	E_Element_State_Long.eWaterReady:;
			IF eReq=E_Request_List.eDissolve THEN;
				eProcess:=E_Element_Process.eDissolving;
			END_IF	
			IF eReq=E_Request_List.eFinish THEN;
				mClearProduction(state:=E_Element_State_Long.eStandby);
			END_IF
	E_Element_State_Long.eReady:;
			IF eReq=E_Request_List.eProduction THEN;
				eProcess:=E_Element_Process.eConnectionToLine;
			END_IF	
			IF eReq=E_Request_List.eFinish THEN;
				mClearProduction(state:=E_Element_State_Long.eStandby);
			END_IF			

	E_Element_State_Long.eProduction:;
			IF eReq=E_Request_List.eDisconnectTank THEN;
				eProcess:=E_Element_Process.eDisconnection;
			END_IF	
			
			IF fbInterConnection_ProL.bAvalableToDisconnect 
			AND m_Production_Run_Pump()
			THEN;
				IF memo_Production_Storage_Mode THEN;
					fb_PumpLine.m_Run(RPM:=stProdParam.stRecipe.FlowRate_Storage);
				ELSE;
					fb_PumpLine.m_Run(RPM:=stProdParam.stRecipe.FlowRate_Production);
				END_IF
				
			ELSE;
				fb_PumpLine.m_Stop();
			END_IF		

	E_Element_State_Long.eEmpty:;
			IF eReq=E_Request_List.eFinish THEN;
				mClearProduction(state:=E_Element_State_Long.eStandby);
			END_IF	

	E_Element_State_Long.eExpired:;
		CASE refElement.eState_Long_Expiered OF
			
			E_Element_State_Long.eProduction:;	
				IF eReq=E_Request_List.eDisconnectTank THEN;
					eProcess:=E_Element_Process.eDisconnection;
				END_IF
				
				IF fbInterConnection_ProL.bAvalableToDisconnect 
				AND m_Production_Run_Pump()
				THEN;
					IF memo_Production_Storage_Mode THEN;
						fb_PumpLine.m_Run(RPM:=stProdParam.stRecipe.FlowRate_Storage);
					ELSE;
						fb_PumpLine.m_Run(RPM:=stProdParam.stRecipe.FlowRate_Production);
					END_IF
					
				ELSE;
					fb_PumpLine.m_Stop();
				END_IF	
		ELSE
			IF eReq=E_Request_List.eFinish THEN;
				mClearProduction(state:=E_Element_State_Long.eStandby);
			END_IF			
		END_CASE
		
END_CASE
END_ACTION

ACTION _aReady_entry:

END_ACTION

ACTION _aReady_exit:
bRun:=TRUE;
bDone:=FALSE;
//bCntrlTemp:=TRUE;
END_ACTION

ACTION _aStart_TriPump_1_active:
bStepDone:=TRUE;
END_ACTION

ACTION _aStart_TriPump_1_entry:
fb_PumpTriBlender.m_Run(RPM:=stProdParam.stRecipe.FlowRate_WaterPushing);
END_ACTION

ACTION _aStart_TriPump_2_active:
bStepDone:=TRUE;
END_ACTION

ACTION _aStart_TriPump_2_entry:
fb_PumpTriBlender.m_Run(RPM:=stProdParam.stRecipe.FlowRate_WaterPushing);
END_ACTION

ACTION _aStart_TriPump_3_active:
bStepDone:=TRUE;
END_ACTION

ACTION _aStart_TriPump_3_entry:
fb_PumpTriBlender.m_Run(RPM:=stProdParam.stRecipe.FlowRate_WaterPushing);
memo_Tank_Level_start:=ref_fbTankSensors.act_Volume;
END_ACTION

ACTION _aState_Update_01_entry:
refState_Long:=E_Element_State_Long.eNotClean;
END_ACTION

ACTION _aState_Update_02_entry:
refState_Long:=E_Element_State_Long.eWaterReady;
END_ACTION

ACTION _aState_Update_03_entry:
refState_Long:=E_Element_State_Long.eReady;
END_ACTION

ACTION _aState_Update_04_entry:
refState_Long:=E_Element_State_Long.eProduction;
END_ACTION

ACTION _aState_Update_05_entry:
refState_Long:=E_Element_State_Long.eReady;
END_ACTION

ACTION _aStop_TriPump_1_active:
bStepDone:=TRUE;
END_ACTION

ACTION _aStop_TriPump_1_entry:
fb_PumpTriBlender.m_Stop();
END_ACTION

ACTION _aStop_TriPump_2_active:
bStepDone:=TRUE;
END_ACTION

ACTION _aStop_TriPump_2_entry:
fb_PumpTriBlender.m_Stop();
END_ACTION

ACTION _aStop_TriPump_3_active:
bStepDone:=TRUE;
END_ACTION

ACTION _aStop_TriPump_3_entry:
fb_PumpTriBlender.m_Stop();
END_ACTION

ACTION _aTank_Drain_active:
bStepDone:=FALSE;
IF fbTarget.m_CheckStatus(eReqStatus:=E_Tank_Target.eDrain) THEN;
	bTON_Active:=TRUE;
	
ELSIF Tank_Drain.t>=T#3S THEN; // max time to detect drain open
	bStepDone:=TRUE;
END_IF
IF Call_TON.Q THEN
	bStepDone:=TRUE;
END_IF
END_ACTION

ACTION _aTank_Drain_entry:
fbTarget.m_Run(eReqProc:=E_Tank_Target.eDrain);
bTON_Active:=FALSE;
END_ACTION

ACTION _aTank_Open_active:
bStepDone:=FALSE;
IF fbTarget.m_CheckStatus(eReqStatus:=E_Tank_Target.eOpen) THEN;
	bTON_Active:=TRUE;
END_IF
IF Call_TON.Q THEN
	bStepDone:=TRUE;
END_IF
END_ACTION

ACTION _aTank_Open_entry:
fbTarget.m_Run(eReqProc:=E_Tank_Target.eOpen);
bTON_Active:=FALSE;
END_ACTION

ACTION _aWater_Fill_active:
bStepDone:=FALSE;
IF TRUE 
AND TRUE//Reserved for tank level from recipe
//AND ref_fbTankSensors.get_stTankLevel().rTankLevel>=stProdParam.stRecipe.arr_Component[1].rWeight
AND fbTarget.stTankLevel.rTankLevel>=stProdParam.stRecipe.arr_Component[1].rWeight
THEN;
	bStepDone:=TRUE;
	
//temp overweight protection
ELSIF stT3_Sens.rTankLevel+stT4_Sens.rTankLevel>1000 THEN;
	bStepDone:=TRUE;
	
ELSIF bRunOffline 
AND Water_Fill.t>=T#10S
THEN
	bStepDone:=TRUE;
END_IF
END_ACTION

ACTION act_Call_Interface:
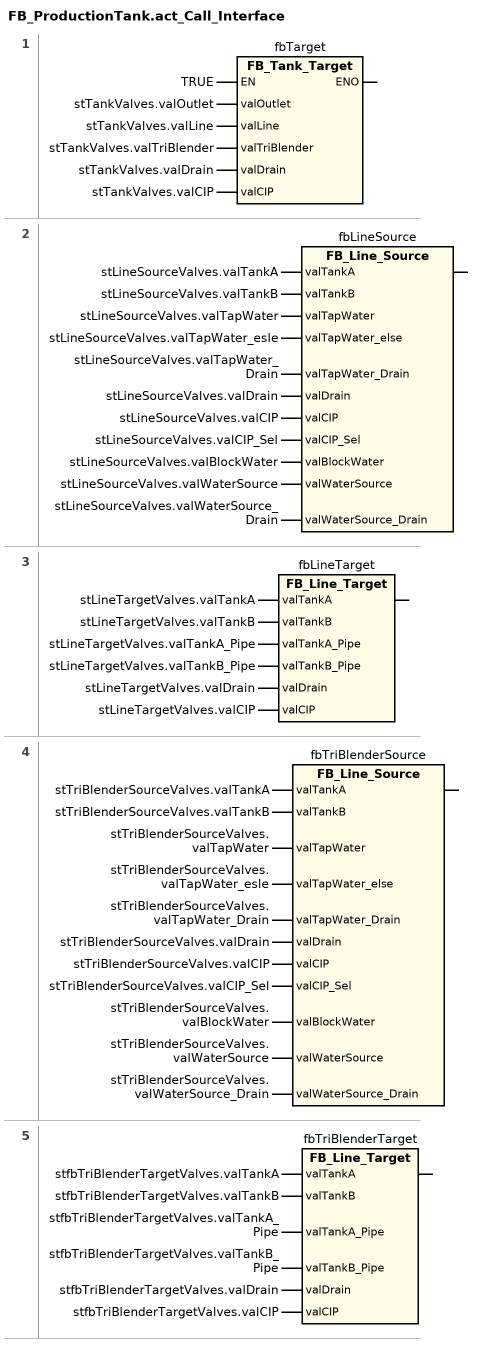
// NETWORK 1
fbTarget(
    valOutlet := stTankValves.valOutlet,
    valLine := stTankValves.valLine,
    valTriBlender := stTankValves.valTriBlender,
    valDrain := stTankValves.valDrain,
    valCIP := stTankValves.valCIP); // FB_Tank_Target

// NETWORK 2
fbLineSource(
    valTankA := stLineSourceValves.valTankA,
    valTankB := stLineSourceValves.valTankB,
    valTapWater := stLineSourceValves.valTapWater,
    valTapWater_else := stLineSourceValves.valTapWater_esle,
    valTapWater_Drain := stLineSourceValves.valTapWater_Drain,
    valDrain := stLineSourceValves.valDrain,
    valCIP := stLineSourceValves.valCIP,
    valCIP_Sel := stLineSourceValves.valCIP_Sel,
    valBlockWater := stLineSourceValves.valBlockWater,
    valWaterSource := stLineSourceValves.valWaterSource,
    valWaterSource_Drain := stLineSourceValves.valWaterSource_Drain); // FB_Line_Source

// NETWORK 3
fbLineTarget(
    valTankA := stLineTargetValves.valTankA,
    valTankB := stLineTargetValves.valTankB,
    valTankA_Pipe := stLineTargetValves.valTankA_Pipe,
    valTankB_Pipe := stLineTargetValves.valTankB_Pipe,
    valDrain := stLineTargetValves.valDrain,
    valCIP := stLineTargetValves.valCIP); // FB_Line_Target

// NETWORK 4
fbTriBlenderSource(
    valTankA := stTriBlenderSourceValves.valTankA,
    valTankB := stTriBlenderSourceValves.valTankB,
    valTapWater := stTriBlenderSourceValves.valTapWater,
    valTapWater_else := stTriBlenderSourceValves.valTapWater_esle,
    valTapWater_Drain := stTriBlenderSourceValves.valTapWater_Drain,
    valDrain := stTriBlenderSourceValves.valDrain,
    valCIP := stTriBlenderSourceValves.valCIP,
    valCIP_Sel := stTriBlenderSourceValves.valCIP_Sel,
    valBlockWater := stTriBlenderSourceValves.valBlockWater,
    valWaterSource := stTriBlenderSourceValves.valWaterSource,
    valWaterSource_Drain := stTriBlenderSourceValves.valWaterSource_Drain); // FB_Line_Source

// NETWORK 5
fbTriBlenderTarget(
    valTankA := stfbTriBlenderTargetValves.valTankA,
    valTankB := stfbTriBlenderTargetValves.valTankB,
    valTankA_Pipe := stfbTriBlenderTargetValves.valTankA_Pipe,
    valTankB_Pipe := stfbTriBlenderTargetValves.valTankB_Pipe,
    valDrain := stfbTriBlenderTargetValves.valDrain,
    valCIP := stfbTriBlenderTargetValves.valCIP); // FB_Line_Target

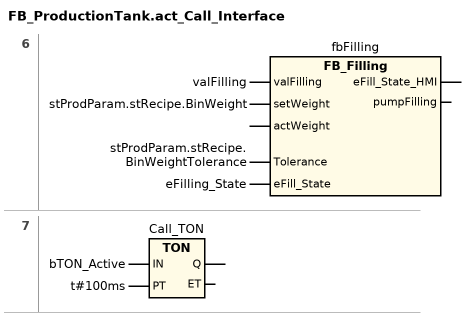
// NETWORK 6
fbFilling(
    valFilling := valFilling,
    setWeight := stProdParam.stRecipe.BinWeight,
    Tolerance := stProdParam.stRecipe.BinWeightTolerance,
    eFill_State := eFilling_State); // FB_Filling

// NETWORK 7
Call_TON(IN := bTON_Active, PT := t#100ms); // TON
END_ACTION

ACTION act_ExpirationTime:
IF stProdParam.eStatus=E_Prod_Status.Active 
THEN;
	refElement.m_Set_ExpirationDuration(eExTime_set:=E_ExTime.eProduct, setTime:=stProdParam.stRecipe.ExpirationTime);
	refElement.m_Set_ExpirationDuration(eExTime_set:=E_ExTime.eWater, setTime:=stProdParam.stRecipe.ExpirationTime_Water);
END_IF


(*
IF stProdParam.eStatus=E_Prod_Status.Active 
AND refElement.State>=E_Element_State_Long.eWaterReady
THEN;
	IF refElement.memoDissolving_active 
	//OR eStatus>=E_Element_State_Long.eReady
	THEN
		refElement.ExpirationTime:=stProdParam.stRecipe.ExpirationTime;
	ELSE;
		refElement.ExpirationTime:=stProdParam.stRecipe.ExpirationTime_Water;
	END_IF
	
ELSE;
	refElement.ExpirationTime:=ExDuration_Default;
END_IF
*)
END_ACTION

ACTION act_Filling:


IF TRUE 
AND bReady
AND refElement.eState_Long=E_Element_State_Long.eProduction
AND TRUE
AND TRUE
THEN;
	CASE pFilling_State OF 
		E_Filling_State.eNot_Ready:;
				pFilling_State:=E_Filling_State.eReady_ToFill;
				
		E_Filling_State.eReady_ToFill:;
				//
		E_Filling_State.eFilling_InProcess:;
				//
		
	END_CASE
ELSE;
	pFilling_State:=E_Filling_State.eNot_Ready;
END_IF

refElement.pFilling_State:=pFilling_State;

(*
IF fbInterConnection_ProL.bActive THEN;
	IF trn_Tank_Marinade THEN;
		fbElement[E_Element_List.eLine_Marinada].pFilling_State:=pFilling_State;
	ELSIF trn_Tank_Color THEN;
		fbElement[E_Element_List.eLine_Color].pFilling_State:=pFilling_State;
	END_IF	
END_IF
*)
END_ACTION

ACTION act_GetReference:
m_Set_SFCFlags_Reference();
refElement REF= fbElement[eElementID];
refState_Long REF= fbElement[eElementID].eState_Long;
//stPis_FillWater REF= stPis[valFillWater];
//stPis_FillWaterDrain REF= stPis[valFillWaterDrain];
//stPis_DrainTapWater REF= stPis[valDrainTapWater];

ref_fbTankSensors REF= g_Data.arrTanksSens[eTank_Name];
stTank_Level:=ref_fbTankSensors.get_stTankLevel();
fbTarget.set_TankLevel(set_stTankLevel:=stTank_Level);

stPis_CWIn REF= stPis[valCW_In];
stPis_CWOut	 REF= stPis[valCW_Out];

eStatus:=refState_Long;

//bRunCIP :=g_Data.b_CIP_Run;
bRunCIP := g_Data.fbElement[eElementID].m_Get_InterConnection() = E_InterConnection.ConnToCIP;
(*
stPis_Outlet		REF= g_Piston.stPis[valOutlet];
stPis_Line			REF= g_Piston.stPis[valOutlet];
stPis_TriBlender	REF= g_Piston.stPis[valOutlet];
stPis_Drain			REF= g_Piston.stPis[valOutlet];
stPis_CIP			REF= g_Piston.stPis[valOutlet];
*)
END_ACTION

ACTION act_Oper:
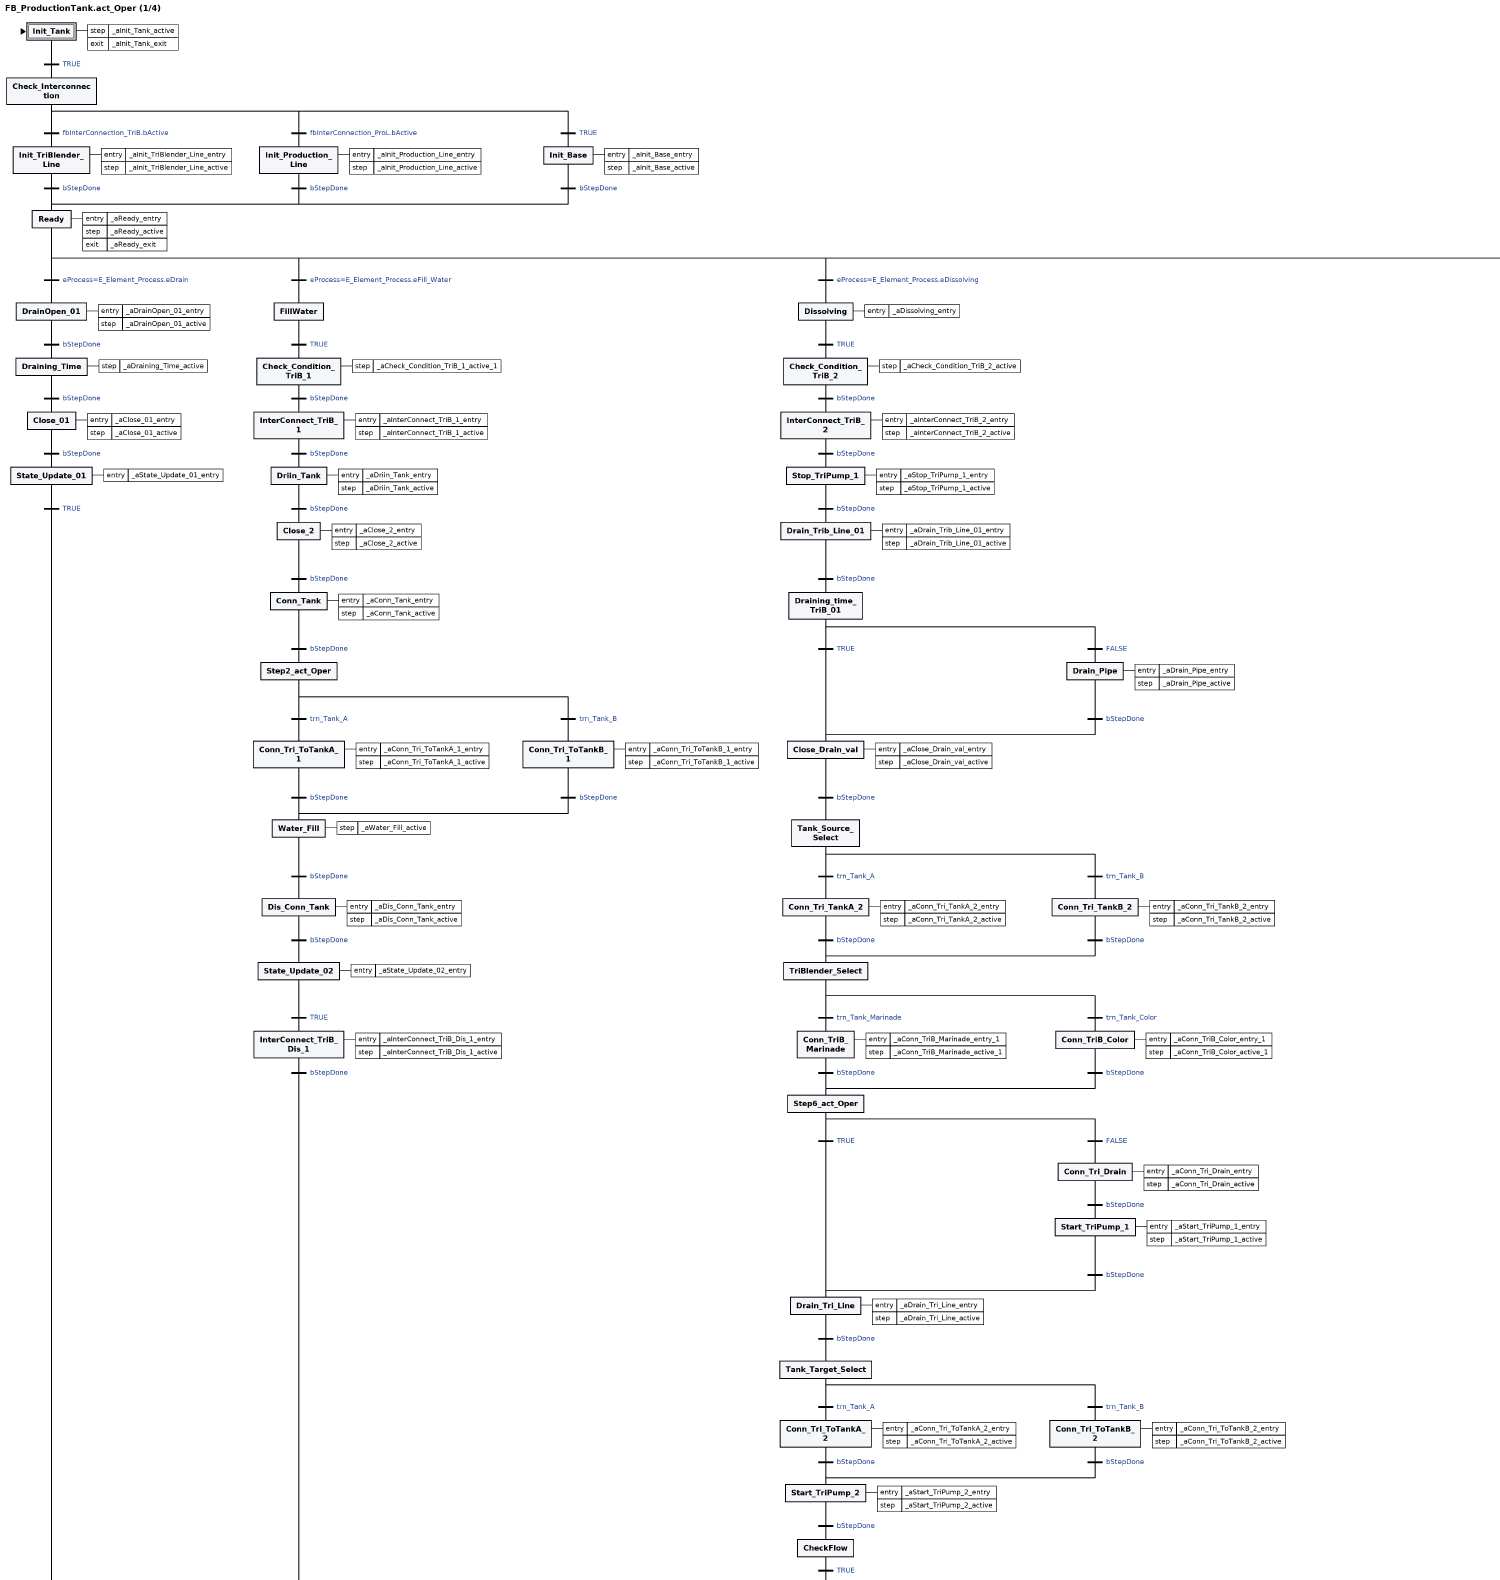
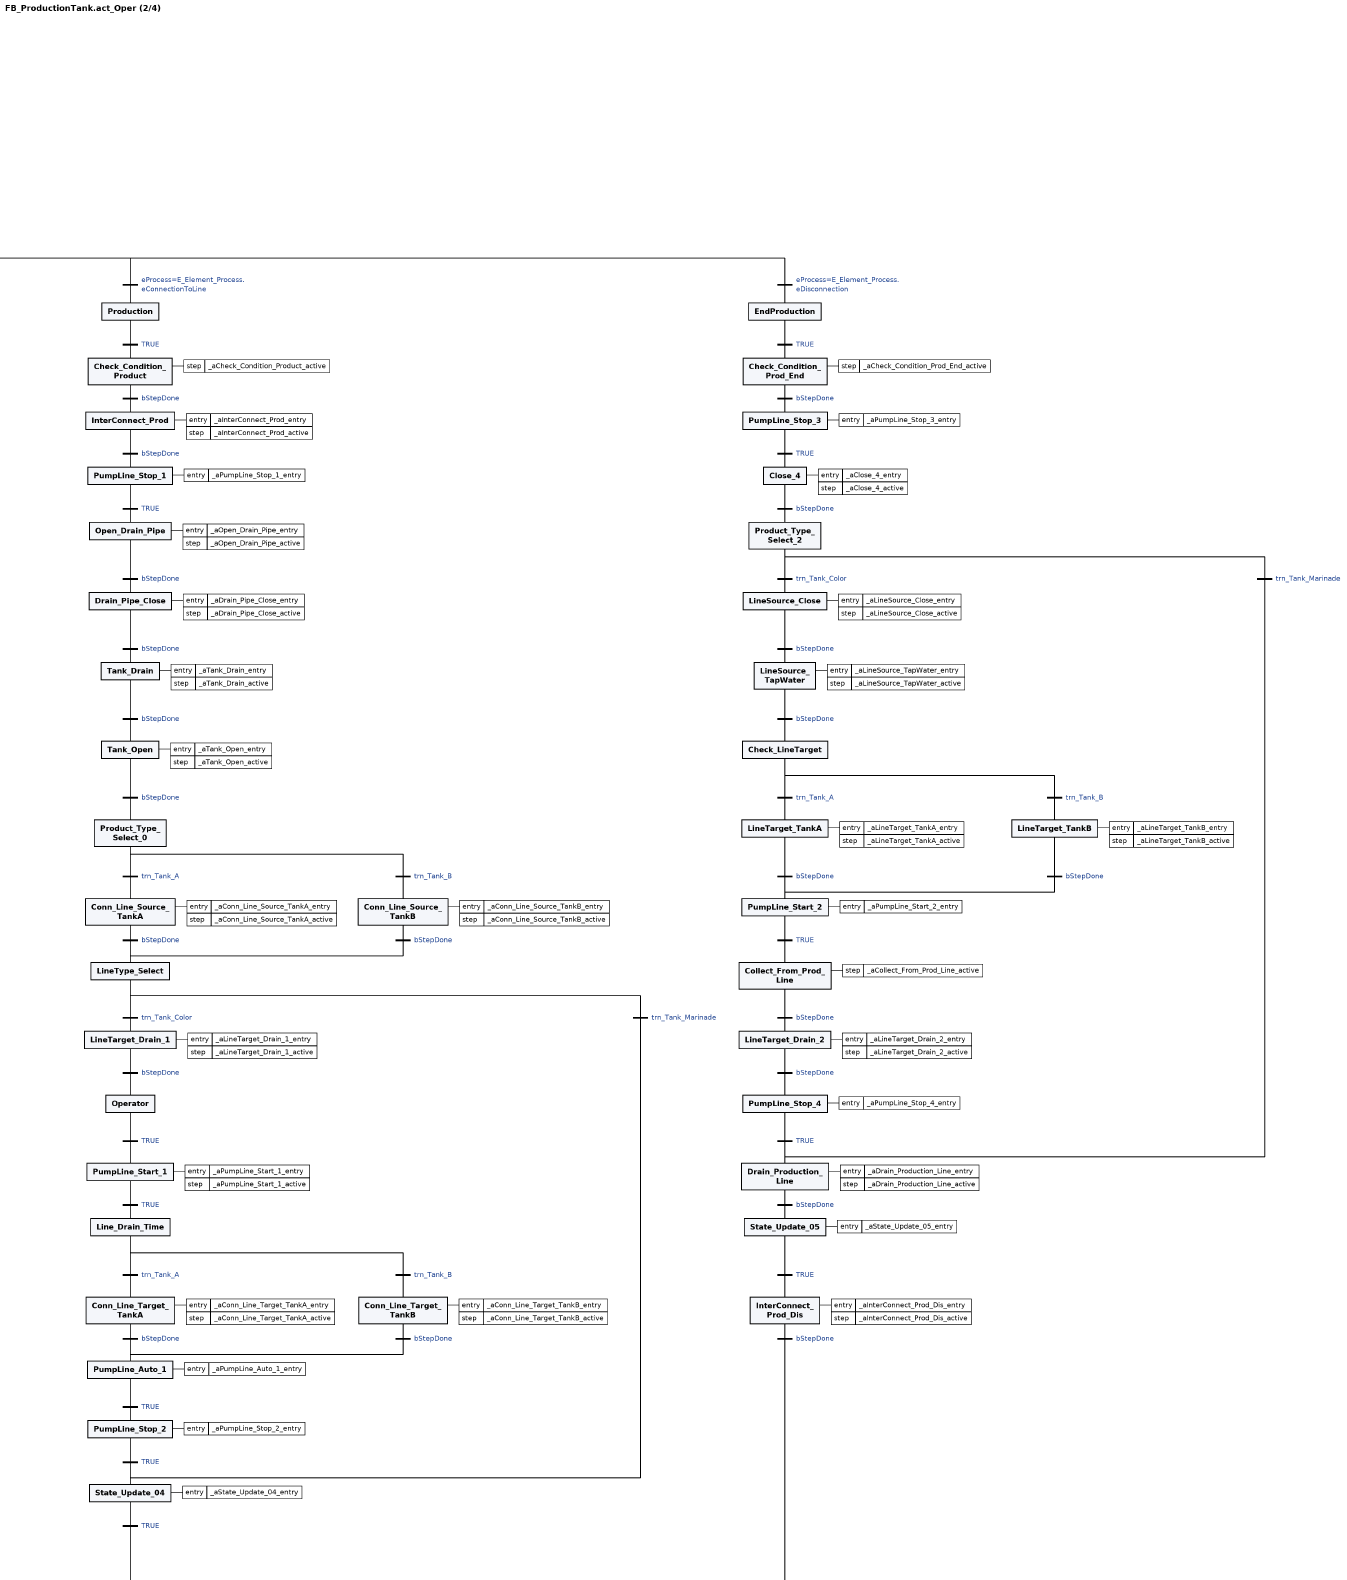
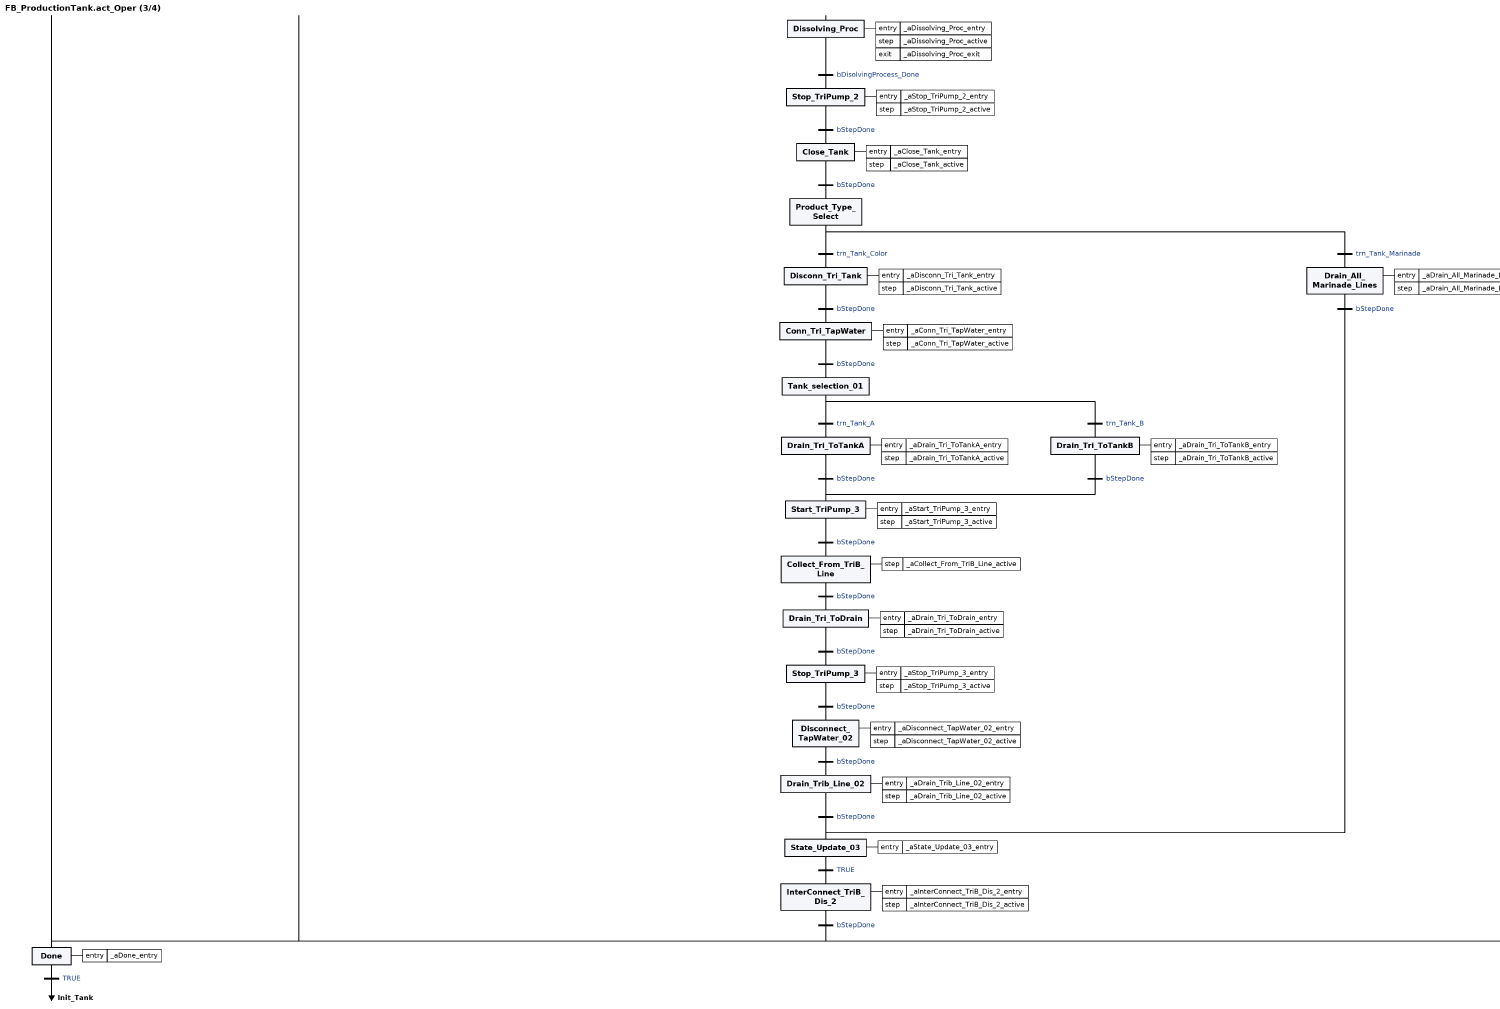
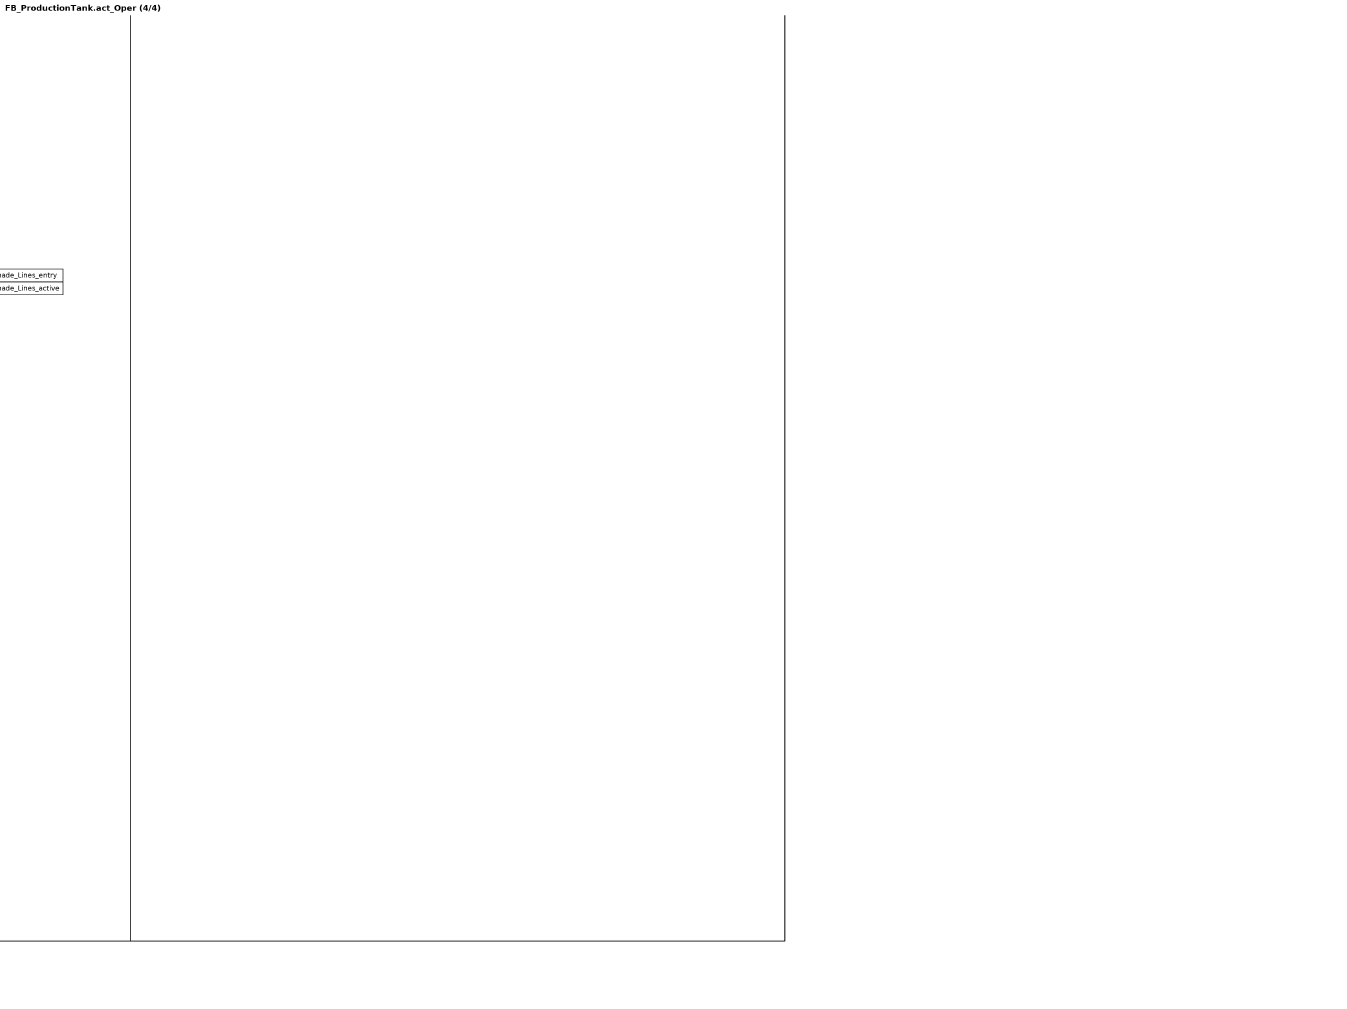
INITIAL_STEP Init_Tank:
    _aInit_Tank_active(N);  // step action
    _aInit_Tank_exit(P0);  // exit action
END_STEP
TRANSITION FROM Init_Tank TO Check_Interconnection
    := TRUE;
END_TRANSITION
STEP Check_Interconnection:
END_STEP
TRANSITION FROM Check_Interconnection TO Init_TriBlender_Line
    := fbInterConnection_TriB.bActive;
END_TRANSITION
STEP Init_TriBlender_Line:
    _aInit_TriBlender_Line_entry(P1);  // entry action
    _aInit_TriBlender_Line_active(N);  // step action
END_STEP
TRANSITION FROM Init_TriBlender_Line TO Ready
    := bStepDone;
END_TRANSITION
TRANSITION FROM Check_Interconnection TO Init_Production_Line
    := fbInterConnection_ProL.bActive;
END_TRANSITION
STEP Init_Production_Line:
    _aInit_Production_Line_entry(P1);  // entry action
    _aInit_Production_Line_active(N);  // step action
END_STEP
TRANSITION FROM Init_Production_Line TO Ready
    := bStepDone;
END_TRANSITION
TRANSITION FROM Check_Interconnection TO Init_Base
    := TRUE;
END_TRANSITION
STEP Init_Base:
    _aInit_Base_entry(P1);  // entry action
    _aInit_Base_active(N);  // step action
END_STEP
TRANSITION FROM Init_Base TO Ready
    := bStepDone;
END_TRANSITION
STEP Ready:
    _aReady_entry(P1);  // entry action
    _aReady_active(N);  // step action
    _aReady_exit(P0);  // exit action
END_STEP
TRANSITION FROM Ready TO DrainOpen_01
    := eProcess=E_Element_Process.eDrain;
END_TRANSITION
STEP DrainOpen_01:  // min time T#2s
    _aDrainOpen_01_entry(P1);  // entry action
    _aDrainOpen_01_active(N);  // step action
END_STEP
TRANSITION FROM DrainOpen_01 TO Draining_Time
    := bStepDone;
END_TRANSITION
STEP Draining_Time:  // min time T#2s
    _aDraining_Time_active(N);  // step action
END_STEP
TRANSITION FROM Draining_Time TO Close_01
    := bStepDone;
END_TRANSITION
STEP Close_01:  // min time T#2s
    _aClose_01_entry(P1);  // entry action
    _aClose_01_active(N);  // step action
END_STEP
TRANSITION FROM Close_01 TO State_Update_01
    := bStepDone;
END_TRANSITION
STEP State_Update_01:
    _aState_Update_01_entry(P1);  // entry action
END_STEP
TRANSITION FROM State_Update_01 TO Done
    := TRUE;
END_TRANSITION
TRANSITION FROM Ready TO FillWater
    := eProcess=E_Element_Process.eFill_Water;
END_TRANSITION
STEP FillWater:
END_STEP
TRANSITION FROM FillWater TO Check_Condition_TriB_1
    := TRUE;
END_TRANSITION
STEP Check_Condition_TriB_1:
    _aCheck_Condition_TriB_1_active_1(N);  // step action
END_STEP
TRANSITION FROM Check_Condition_TriB_1 TO InterConnect_TriB_1
    := bStepDone;
END_TRANSITION
STEP InterConnect_TriB_1:
    _aInterConnect_TriB_1_entry(P1);  // entry action
    _aInterConnect_TriB_1_active(N);  // step action
END_STEP
TRANSITION FROM InterConnect_TriB_1 TO Driin_Tank
    := bStepDone;
END_TRANSITION
STEP Driin_Tank:  // min time t#2s
    _aDriin_Tank_entry(P1);  // entry action
    _aDriin_Tank_active(N);  // step action
END_STEP
TRANSITION FROM Driin_Tank TO Close_2
    := bStepDone;
END_TRANSITION
STEP Close_2:  // min time t#2s
    _aClose_2_entry(P1);  // entry action
    _aClose_2_active(N);  // step action
END_STEP
TRANSITION FROM Close_2 TO Conn_Tank
    := bStepDone;
END_TRANSITION
STEP Conn_Tank:  // min time t#2s
    _aConn_Tank_entry(P1);  // entry action
    _aConn_Tank_active(N);  // step action
END_STEP
TRANSITION FROM Conn_Tank TO Step2_act_Oper
    := bStepDone;
END_TRANSITION
STEP Step2_act_Oper:
END_STEP
TRANSITION FROM Step2_act_Oper TO Conn_Tri_ToTankA_1
    := trn_Tank_A;
END_TRANSITION
STEP Conn_Tri_ToTankA_1:
    _aConn_Tri_ToTankA_1_entry(P1);  // entry action
    _aConn_Tri_ToTankA_1_active(N);  // step action
END_STEP
TRANSITION FROM Conn_Tri_ToTankA_1 TO Water_Fill
    := bStepDone;
END_TRANSITION
TRANSITION FROM Step2_act_Oper TO Conn_Tri_ToTankB_1
    := trn_Tank_B;
END_TRANSITION
STEP Conn_Tri_ToTankB_1:
    _aConn_Tri_ToTankB_1_entry(P1);  // entry action
    _aConn_Tri_ToTankB_1_active(N);  // step action
END_STEP
TRANSITION FROM Conn_Tri_ToTankB_1 TO Water_Fill
    := bStepDone;
END_TRANSITION
STEP Water_Fill:  // min time t#2s
    _aWater_Fill_active(N);  // step action
END_STEP
TRANSITION FROM Water_Fill TO Dis_Conn_Tank
    := bStepDone;
END_TRANSITION
STEP Dis_Conn_Tank:  // min time t#2s
    _aDis_Conn_Tank_entry(P1);  // entry action
    _aDis_Conn_Tank_active(N);  // step action
END_STEP
TRANSITION FROM Dis_Conn_Tank TO State_Update_02
    := bStepDone;
END_TRANSITION
STEP State_Update_02:  // min time t#2s
    _aState_Update_02_entry(P1);  // entry action
END_STEP
TRANSITION FROM State_Update_02 TO InterConnect_TriB_Dis_1
    := TRUE;
END_TRANSITION
STEP InterConnect_TriB_Dis_1:
    _aInterConnect_TriB_Dis_1_entry(P1);  // entry action
    _aInterConnect_TriB_Dis_1_active(N);  // step action
END_STEP
TRANSITION FROM InterConnect_TriB_Dis_1 TO Done
    := bStepDone;
END_TRANSITION
TRANSITION FROM Ready TO Dissolving
    := eProcess=E_Element_Process.eDissolving;
END_TRANSITION
STEP Dissolving:
    _aDissolving_entry(P1);  // entry action
END_STEP
TRANSITION FROM Dissolving TO Check_Condition_TriB_2
    := TRUE;
END_TRANSITION
STEP Check_Condition_TriB_2:
    _aCheck_Condition_TriB_2_active(N);  // step action
END_STEP
TRANSITION FROM Check_Condition_TriB_2 TO InterConnect_TriB_2
    := bStepDone;
END_TRANSITION
STEP InterConnect_TriB_2:
    _aInterConnect_TriB_2_entry(P1);  // entry action
    _aInterConnect_TriB_2_active(N);  // step action
END_STEP
TRANSITION FROM InterConnect_TriB_2 TO Stop_TriPump_1
    := bStepDone;
END_TRANSITION
STEP Stop_TriPump_1:
    _aStop_TriPump_1_entry(P1);  // entry action
    _aStop_TriPump_1_active(N);  // step action
END_STEP
TRANSITION FROM Stop_TriPump_1 TO Drain_Trib_Line_01
    := bStepDone;
END_TRANSITION
STEP Drain_Trib_Line_01:
    _aDrain_Trib_Line_01_entry(P1);  // entry action
    _aDrain_Trib_Line_01_active(N);  // step action
END_STEP
TRANSITION FROM Drain_Trib_Line_01 TO Draining_time_TriB_01
    := bStepDone;
END_TRANSITION
STEP Draining_time_TriB_01:  // min time T#10s
END_STEP
TRANSITION FROM Draining_time_TriB_01 TO Close_Drain_val
    := TRUE;
END_TRANSITION
TRANSITION FROM Draining_time_TriB_01 TO Drain_Pipe
    := FALSE;
END_TRANSITION
STEP Drain_Pipe:  // min time T#2s
    _aDrain_Pipe_entry(P1);  // entry action
    _aDrain_Pipe_active(N);  // step action
END_STEP
TRANSITION FROM Drain_Pipe TO Close_Drain_val
    := bStepDone;
END_TRANSITION
STEP Close_Drain_val:
    _aClose_Drain_val_entry(P1);  // entry action
    _aClose_Drain_val_active(N);  // step action
END_STEP
TRANSITION FROM Close_Drain_val TO Tank_Source_Select
    := bStepDone;
END_TRANSITION
STEP Tank_Source_Select:
END_STEP
TRANSITION FROM Tank_Source_Select TO Conn_Tri_TankA_2
    := trn_Tank_A;
END_TRANSITION
STEP Conn_Tri_TankA_2:
    _aConn_Tri_TankA_2_entry(P1);  // entry action
    _aConn_Tri_TankA_2_active(N);  // step action
END_STEP
TRANSITION FROM Conn_Tri_TankA_2 TO TriBlender_Select
    := bStepDone;
END_TRANSITION
TRANSITION FROM Tank_Source_Select TO Conn_Tri_TankB_2
    := trn_Tank_B;
END_TRANSITION
STEP Conn_Tri_TankB_2:
    _aConn_Tri_TankB_2_entry(P1);  // entry action
    _aConn_Tri_TankB_2_active(N);  // step action
END_STEP
TRANSITION FROM Conn_Tri_TankB_2 TO TriBlender_Select
    := bStepDone;
END_TRANSITION
STEP TriBlender_Select:
END_STEP
TRANSITION FROM TriBlender_Select TO Conn_TriB_Marinade
    := trn_Tank_Marinade;
END_TRANSITION
STEP Conn_TriB_Marinade:
    _aConn_TriB_Marinade_entry_1(P1);  // entry action
    _aConn_TriB_Marinade_active_1(N);  // step action
END_STEP
TRANSITION FROM Conn_TriB_Marinade TO Step6_act_Oper
    := bStepDone;
END_TRANSITION
TRANSITION FROM TriBlender_Select TO Conn_TriB_Color
    := trn_Tank_Color;
END_TRANSITION
STEP Conn_TriB_Color:
    _aConn_TriB_Color_entry_1(P1);  // entry action
    _aConn_TriB_Color_active_1(N);  // step action
END_STEP
TRANSITION FROM Conn_TriB_Color TO Step6_act_Oper
    := bStepDone;
END_TRANSITION
STEP Step6_act_Oper:
END_STEP
TRANSITION FROM Step6_act_Oper TO Drain_Tri_Line
    := TRUE;
END_TRANSITION
TRANSITION FROM Step6_act_Oper TO Conn_Tri_Drain
    := FALSE;
END_TRANSITION
STEP Conn_Tri_Drain:
    _aConn_Tri_Drain_entry(P1);  // entry action
    _aConn_Tri_Drain_active(N);  // step action
END_STEP
TRANSITION FROM Conn_Tri_Drain TO Start_TriPump_1
    := bStepDone;
END_TRANSITION
STEP Start_TriPump_1:
    _aStart_TriPump_1_entry(P1);  // entry action
    _aStart_TriPump_1_active(N);  // step action
END_STEP
TRANSITION FROM Start_TriPump_1 TO Drain_Tri_Line
    := bStepDone;
END_TRANSITION
STEP Drain_Tri_Line:  // min time T#10s
    _aDrain_Tri_Line_entry(P1);  // entry action
    _aDrain_Tri_Line_active(N);  // step action
END_STEP
TRANSITION FROM Drain_Tri_Line TO Tank_Target_Select
    := bStepDone;
END_TRANSITION
STEP Tank_Target_Select:
END_STEP
TRANSITION FROM Tank_Target_Select TO Conn_Tri_ToTankA_2
    := trn_Tank_A;
END_TRANSITION
STEP Conn_Tri_ToTankA_2:
    _aConn_Tri_ToTankA_2_entry(P1);  // entry action
    _aConn_Tri_ToTankA_2_active(N);  // step action
END_STEP
TRANSITION FROM Conn_Tri_ToTankA_2 TO Start_TriPump_2
    := bStepDone;
END_TRANSITION
TRANSITION FROM Tank_Target_Select TO Conn_Tri_ToTankB_2
    := trn_Tank_B;
END_TRANSITION
STEP Conn_Tri_ToTankB_2:
    _aConn_Tri_ToTankB_2_entry(P1);  // entry action
    _aConn_Tri_ToTankB_2_active(N);  // step action
END_STEP
TRANSITION FROM Conn_Tri_ToTankB_2 TO Start_TriPump_2
    := bStepDone;
END_TRANSITION
STEP Start_TriPump_2:
    _aStart_TriPump_2_entry(P1);  // entry action
    _aStart_TriPump_2_active(N);  // step action
END_STEP
TRANSITION FROM Start_TriPump_2 TO CheckFlow
    := bStepDone;
END_TRANSITION
STEP CheckFlow:  // min time t#20s
END_STEP
TRANSITION FROM CheckFlow TO Dissolving_Proc
    := TRUE;
END_TRANSITION
STEP Dissolving_Proc:
    _aDissolving_Proc_entry(P1);  // entry action
    _aDissolving_Proc_active(N);  // step action
    _aDissolving_Proc_exit(P0);  // exit action
END_STEP
TRANSITION FROM Dissolving_Proc TO Stop_TriPump_2
    := bDisolvingProcess_Done;
END_TRANSITION
STEP Stop_TriPump_2:  // min time T#5s
    _aStop_TriPump_2_entry(P1);  // entry action
    _aStop_TriPump_2_active(N);  // step action
END_STEP
TRANSITION FROM Stop_TriPump_2 TO Close_Tank
    := bStepDone;
END_TRANSITION
STEP Close_Tank:
    _aClose_Tank_entry(P1);  // entry action
    _aClose_Tank_active(N);  // step action
END_STEP
TRANSITION FROM Close_Tank TO Product_Type_Select
    := bStepDone;
END_TRANSITION
STEP Product_Type_Select:
END_STEP
TRANSITION FROM Product_Type_Select TO Disconn_Tri_Tank
    := trn_Tank_Color;
END_TRANSITION
STEP Disconn_Tri_Tank:  // min time t#100ms
    _aDisconn_Tri_Tank_entry(P1);  // entry action
    _aDisconn_Tri_Tank_active(N);  // step action
END_STEP
TRANSITION FROM Disconn_Tri_Tank TO Conn_Tri_TapWater
    := bStepDone;
END_TRANSITION
STEP Conn_Tri_TapWater:  // min time T#5s
    _aConn_Tri_TapWater_entry(P1);  // entry action
    _aConn_Tri_TapWater_active(N);  // step action
END_STEP
TRANSITION FROM Conn_Tri_TapWater TO Tank_selection_01
    := bStepDone;
END_TRANSITION
STEP Tank_selection_01:
END_STEP
TRANSITION FROM Tank_selection_01 TO Drain_Tri_ToTankA
    := trn_Tank_A;
END_TRANSITION
STEP Drain_Tri_ToTankA:  // min time t#100ms
    _aDrain_Tri_ToTankA_entry(P1);  // entry action
    _aDrain_Tri_ToTankA_active(N);  // step action
END_STEP
TRANSITION FROM Drain_Tri_ToTankA TO Start_TriPump_3
    := bStepDone;
END_TRANSITION
TRANSITION FROM Tank_selection_01 TO Drain_Tri_ToTankB
    := trn_Tank_B;
END_TRANSITION
STEP Drain_Tri_ToTankB:  // min time t#100ms
    _aDrain_Tri_ToTankB_entry(P1);  // entry action
    _aDrain_Tri_ToTankB_active(N);  // step action
END_STEP
TRANSITION FROM Drain_Tri_ToTankB TO Start_TriPump_3
    := bStepDone;
END_TRANSITION
STEP Start_TriPump_3:
    _aStart_TriPump_3_entry(P1);  // entry action
    _aStart_TriPump_3_active(N);  // step action
END_STEP
TRANSITION FROM Start_TriPump_3 TO Collect_From_TriB_Line
    := bStepDone;
END_TRANSITION
STEP Collect_From_TriB_Line:
    _aCollect_From_TriB_Line_active(N);  // step action
END_STEP
TRANSITION FROM Collect_From_TriB_Line TO Drain_Tri_ToDrain
    := bStepDone;
END_TRANSITION
STEP Drain_Tri_ToDrain:  // min time T#25s
    _aDrain_Tri_ToDrain_entry(P1);  // entry action
    _aDrain_Tri_ToDrain_active(N);  // step action
END_STEP
TRANSITION FROM Drain_Tri_ToDrain TO Stop_TriPump_3
    := bStepDone;
END_TRANSITION
STEP Stop_TriPump_3:
    _aStop_TriPump_3_entry(P1);  // entry action
    _aStop_TriPump_3_active(N);  // step action
END_STEP
TRANSITION FROM Stop_TriPump_3 TO Disconnect_TapWater_02
    := bStepDone;
END_TRANSITION
STEP Disconnect_TapWater_02:
    _aDisconnect_TapWater_02_entry(P1);  // entry action
    _aDisconnect_TapWater_02_active(N);  // step action
END_STEP
TRANSITION FROM Disconnect_TapWater_02 TO Drain_Trib_Line_02
    := bStepDone;
END_TRANSITION
STEP Drain_Trib_Line_02:  // min time T#10s
    _aDrain_Trib_Line_02_entry(P1);  // entry action
    _aDrain_Trib_Line_02_active(N);  // step action
END_STEP
TRANSITION FROM Drain_Trib_Line_02 TO State_Update_03
    := bStepDone;
END_TRANSITION
TRANSITION FROM Product_Type_Select TO Drain_All_Marinade_Lines
    := trn_Tank_Marinade;
END_TRANSITION
STEP Drain_All_Marinade_Lines:
    _aDrain_All_Marinade_Lines_entry(P1);  // entry action
    _aDrain_All_Marinade_Lines_active(N);  // step action
END_STEP
TRANSITION FROM Drain_All_Marinade_Lines TO State_Update_03
    := bStepDone;
END_TRANSITION
STEP State_Update_03:
    _aState_Update_03_entry(P1);  // entry action
END_STEP
TRANSITION FROM State_Update_03 TO InterConnect_TriB_Dis_2
    := TRUE;
END_TRANSITION
STEP InterConnect_TriB_Dis_2:
    _aInterConnect_TriB_Dis_2_entry(P1);  // entry action
    _aInterConnect_TriB_Dis_2_active(N);  // step action
END_STEP
TRANSITION FROM InterConnect_TriB_Dis_2 TO Done
    := bStepDone;
END_TRANSITION
TRANSITION FROM Ready TO Production
    := eProcess=E_Element_Process.eConnectionToLine;
END_TRANSITION
STEP Production:
END_STEP
TRANSITION FROM Production TO Check_Condition_Product
    := TRUE;
END_TRANSITION
STEP Check_Condition_Product:
    _aCheck_Condition_Product_active(N);  // step action
END_STEP
TRANSITION FROM Check_Condition_Product TO InterConnect_Prod
    := bStepDone;
END_TRANSITION
STEP InterConnect_Prod:
    _aInterConnect_Prod_entry(P1);  // entry action
    _aInterConnect_Prod_active(N);  // step action
END_STEP
TRANSITION FROM InterConnect_Prod TO PumpLine_Stop_1
    := bStepDone;
END_TRANSITION
STEP PumpLine_Stop_1:
    _aPumpLine_Stop_1_entry(P1);  // entry action
END_STEP
TRANSITION FROM PumpLine_Stop_1 TO Open_Drain_Pipe
    := TRUE;
END_TRANSITION
STEP Open_Drain_Pipe:  // min time T#5s
    _aOpen_Drain_Pipe_entry(P1);  // entry action
    _aOpen_Drain_Pipe_active(N);  // step action
END_STEP
TRANSITION FROM Open_Drain_Pipe TO Drain_Pipe_Close
    := bStepDone;
END_TRANSITION
STEP Drain_Pipe_Close:
    _aDrain_Pipe_Close_entry(P1);  // entry action
    _aDrain_Pipe_Close_active(N);  // step action
END_STEP
TRANSITION FROM Drain_Pipe_Close TO Tank_Drain
    := bStepDone;
END_TRANSITION
STEP Tank_Drain:  // min time t#2s
    _aTank_Drain_entry(P1);  // entry action
    _aTank_Drain_active(N);  // step action
END_STEP
TRANSITION FROM Tank_Drain TO Tank_Open
    := bStepDone;
END_TRANSITION
STEP Tank_Open:  // min time t#2s
    _aTank_Open_entry(P1);  // entry action
    _aTank_Open_active(N);  // step action
END_STEP
TRANSITION FROM Tank_Open TO Product_Type_Select_0
    := bStepDone;
END_TRANSITION
STEP Product_Type_Select_0:
END_STEP
TRANSITION FROM Product_Type_Select_0 TO Conn_Line_Source_TankA
    := trn_Tank_A;
END_TRANSITION
STEP Conn_Line_Source_TankA:  // min time t#100ms
    _aConn_Line_Source_TankA_entry(P1);  // entry action
    _aConn_Line_Source_TankA_active(N);  // step action
END_STEP
TRANSITION FROM Conn_Line_Source_TankA TO LineType_Select
    := bStepDone;
END_TRANSITION
TRANSITION FROM Product_Type_Select_0 TO Conn_Line_Source_TankB
    := trn_Tank_B;
END_TRANSITION
STEP Conn_Line_Source_TankB:  // min time t#100ms
    _aConn_Line_Source_TankB_entry(P1);  // entry action
    _aConn_Line_Source_TankB_active(N);  // step action
END_STEP
TRANSITION FROM Conn_Line_Source_TankB TO LineType_Select
    := bStepDone;
END_TRANSITION
STEP LineType_Select:
END_STEP
TRANSITION FROM LineType_Select TO LineTarget_Drain_1
    := trn_Tank_Color;
END_TRANSITION
STEP LineTarget_Drain_1:
    _aLineTarget_Drain_1_entry(P1);  // entry action
    _aLineTarget_Drain_1_active(N);  // step action
END_STEP
TRANSITION FROM LineTarget_Drain_1 TO Operator
    := bStepDone;
END_TRANSITION
STEP Operator:
END_STEP
TRANSITION FROM Operator TO PumpLine_Start_1
    := TRUE;
END_TRANSITION
STEP PumpLine_Start_1:
    _aPumpLine_Start_1_entry(P1);  // entry action
    _aPumpLine_Start_1_active(N);  // step action
END_STEP
TRANSITION FROM PumpLine_Start_1 TO Line_Drain_Time
    := TRUE;
END_TRANSITION
STEP Line_Drain_Time:  // min time T#10s
END_STEP
TRANSITION FROM Line_Drain_Time TO Conn_Line_Target_TankA
    := trn_Tank_A;
END_TRANSITION
STEP Conn_Line_Target_TankA:
    _aConn_Line_Target_TankA_entry(P1);  // entry action
    _aConn_Line_Target_TankA_active(N);  // step action
END_STEP
TRANSITION FROM Conn_Line_Target_TankA TO PumpLine_Auto_1
    := bStepDone;
END_TRANSITION
TRANSITION FROM Line_Drain_Time TO Conn_Line_Target_TankB
    := trn_Tank_B;
END_TRANSITION
STEP Conn_Line_Target_TankB:
    _aConn_Line_Target_TankB_entry(P1);  // entry action
    _aConn_Line_Target_TankB_active(N);  // step action
END_STEP
TRANSITION FROM Conn_Line_Target_TankB TO PumpLine_Auto_1
    := bStepDone;
END_TRANSITION
STEP PumpLine_Auto_1:
    _aPumpLine_Auto_1_entry(P1);  // entry action
END_STEP
TRANSITION FROM PumpLine_Auto_1 TO PumpLine_Stop_2
    := TRUE;
END_TRANSITION
STEP PumpLine_Stop_2:
    _aPumpLine_Stop_2_entry(P1);  // entry action
END_STEP
TRANSITION FROM PumpLine_Stop_2 TO State_Update_04
    := TRUE;
END_TRANSITION
TRANSITION FROM LineType_Select TO State_Update_04
    := trn_Tank_Marinade;
END_TRANSITION
STEP State_Update_04:
    _aState_Update_04_entry(P1);  // entry action
END_STEP
TRANSITION FROM State_Update_04 TO Done
    := TRUE;
END_TRANSITION
TRANSITION FROM Ready TO EndProduction
    := eProcess=E_Element_Process.eDisconnection;
END_TRANSITION
STEP EndProduction:
END_STEP
TRANSITION FROM EndProduction TO Check_Condition_Prod_End
    := TRUE;
END_TRANSITION
STEP Check_Condition_Prod_End:
    _aCheck_Condition_Prod_End_active(N);  // step action
END_STEP
TRANSITION FROM Check_Condition_Prod_End TO PumpLine_Stop_3
    := bStepDone;
END_TRANSITION
STEP PumpLine_Stop_3:
    _aPumpLine_Stop_3_entry(P1);  // entry action
END_STEP
TRANSITION FROM PumpLine_Stop_3 TO Close_4
    := TRUE;
END_TRANSITION
STEP Close_4:
    _aClose_4_entry(P1);  // entry action
    _aClose_4_active(N);  // step action
END_STEP
TRANSITION FROM Close_4 TO Product_Type_Select_2
    := bStepDone;
END_TRANSITION
STEP Product_Type_Select_2:
END_STEP
TRANSITION FROM Product_Type_Select_2 TO LineSource_Close
    := trn_Tank_Color;
END_TRANSITION
STEP LineSource_Close:
    _aLineSource_Close_entry(P1);  // entry action
    _aLineSource_Close_active(N);  // step action
END_STEP
TRANSITION FROM LineSource_Close TO LineSource_TapWater
    := bStepDone;
END_TRANSITION
STEP LineSource_TapWater:
    _aLineSource_TapWater_entry(P1);  // entry action
    _aLineSource_TapWater_active(N);  // step action
END_STEP
TRANSITION FROM LineSource_TapWater TO Check_LineTarget
    := bStepDone;
END_TRANSITION
STEP Check_LineTarget:
END_STEP
TRANSITION FROM Check_LineTarget TO LineTarget_TankA
    := trn_Tank_A;
END_TRANSITION
STEP LineTarget_TankA:
    _aLineTarget_TankA_entry(P1);  // entry action
    _aLineTarget_TankA_active(N);  // step action
END_STEP
TRANSITION FROM LineTarget_TankA TO PumpLine_Start_2
    := bStepDone;
END_TRANSITION
TRANSITION FROM Check_LineTarget TO LineTarget_TankB
    := trn_Tank_B;
END_TRANSITION
STEP LineTarget_TankB:
    _aLineTarget_TankB_entry(P1);  // entry action
    _aLineTarget_TankB_active(N);  // step action
END_STEP
TRANSITION FROM LineTarget_TankB TO PumpLine_Start_2
    := bStepDone;
END_TRANSITION
STEP PumpLine_Start_2:
    _aPumpLine_Start_2_entry(P1);  // entry action
END_STEP
TRANSITION FROM PumpLine_Start_2 TO Collect_From_Prod_Line
    := TRUE;
END_TRANSITION
STEP Collect_From_Prod_Line:
    _aCollect_From_Prod_Line_active(N);  // step action
END_STEP
TRANSITION FROM Collect_From_Prod_Line TO LineTarget_Drain_2
    := bStepDone;
END_TRANSITION
STEP LineTarget_Drain_2:  // min time T#25s
    _aLineTarget_Drain_2_entry(P1);  // entry action
    _aLineTarget_Drain_2_active(N);  // step action
END_STEP
TRANSITION FROM LineTarget_Drain_2 TO PumpLine_Stop_4
    := bStepDone;
END_TRANSITION
STEP PumpLine_Stop_4:
    _aPumpLine_Stop_4_entry(P1);  // entry action
END_STEP
TRANSITION FROM PumpLine_Stop_4 TO Drain_Production_Line
    := TRUE;
END_TRANSITION
TRANSITION FROM Product_Type_Select_2 TO Drain_Production_Line
    := trn_Tank_Marinade;
END_TRANSITION
STEP Drain_Production_Line:
    _aDrain_Production_Line_entry(P1);  // entry action
    _aDrain_Production_Line_active(N);  // step action
END_STEP
TRANSITION FROM Drain_Production_Line TO State_Update_05
    := bStepDone;
END_TRANSITION
STEP State_Update_05:
    _aState_Update_05_entry(P1);  // entry action
END_STEP
TRANSITION FROM State_Update_05 TO InterConnect_Prod_Dis
    := TRUE;
END_TRANSITION
STEP InterConnect_Prod_Dis:
    _aInterConnect_Prod_Dis_entry(P1);  // entry action
    _aInterConnect_Prod_Dis_active(N);  // step action
END_STEP
TRANSITION FROM InterConnect_Prod_Dis TO Done
    := bStepDone;
END_TRANSITION
STEP Done:  // min time T#2s
    _aDone_entry(P1);  // entry action
END_STEP
TRANSITION FROM Done TO Init_Tank
    := TRUE;
END_TRANSITION
// branch label Branch11_act_Oper
// branch label Branch3_act_Oper
// branch label Branch10_act_Oper
// branch label Branch1_act_Oper
// branch label Branch7_act_Oper
// branch label Branch9_act_Oper
// branch label Branch2_act_Oper
// branch label Branch8_act_Oper
// branch label Branch4_act_Oper
// branch label Branch5_act_Oper
// branch label Branch14_act_Oper
// branch label Branch6_act_Oper
// branch label Branch12_act_Oper
// branch label Branch0_act_Oper_Tank
END_ACTION

ACTION act_TempCntrl:
CASE eElementID OF 
	E_Element_List.eTank_1:
		//Marinada Tank 1
		st_TempCntrl 	REF=g_ProcControl.arr_stProcCntrl[E_ProcessControl_Name.eMarinTank1_Temp];
		pc_TempCntrl 	REF= g_ProcControl.arr_fbProcCntrl[E_ProcessControl_Name.eMarinTank1_Temp];
		//tolerance
	E_Element_List.eTank_2:
		//Marinada Tank 2
		st_TempCntrl 	REF=g_ProcControl.arr_stProcCntrl[E_ProcessControl_Name.eMarinTank2_Temp];
		pc_TempCntrl 	REF= g_ProcControl.arr_fbProcCntrl[E_ProcessControl_Name.eMarinTank2_Temp];
	E_Element_List.eTank_3:
		//Color Tank 1
		st_TempCntrl 	REF=g_ProcControl.arr_stProcCntrl[E_ProcessControl_Name.eColorTank1_Temp];
		pc_TempCntrl 	REF= g_ProcControl.arr_fbProcCntrl[E_ProcessControl_Name.eColorTank1_Temp];
	E_Element_List.eTank_4:
		//Color Tank 2
		st_TempCntrl 	REF=g_ProcControl.arr_stProcCntrl[E_ProcessControl_Name.eColorTank2_Temp];
		pc_TempCntrl 	REF= g_ProcControl.arr_fbProcCntrl[E_ProcessControl_Name.eColorTank2_Temp];
END_CASE
st_TempCntrl.rValue:=g_AnalogSensor.stAnalogSensor[sens_TankTemp].Value;//sensor
//st_TempCntrl.rValue:=rTest;//sensor test
st_TempCntrl.rSetPoint:=stProdParam.stRecipe.Temperature;//value from recipe
st_TempCntrl.fHystLow:=stProdParam.stRecipe.Temperature-1;
st_TempCntrl.fHystHigh:=stProdParam.stRecipe.Temperature+0.5;
//st_TempCntrl.ToleranceHigh:=5;
//st_TempCntrl.ToleravceLow:=-55;



bCntrlTemp:=stProdParam.eStatus=E_Prod_Status.Active
AND eStatus>=E_Element_State_Long.eWaterReady;

IF bCntrlTemp AND NOT bRunCIP THEN
	//pc_TempCntrl.mRun_Hyst();
	pc_TempCntrl(stProcessControl:=st_TempCntrl);
	
 	IF TRUE 
	AND (NOT st_TempCntrl.bHystOut)
	AND  stPis_CWOut.st_Close
	THEN
		stPis_CWOut.req_Open:=TRUE;
		
	ELSIF (st_TempCntrl.bHystOut)
	AND stPis_CWOut.st_Open THEN;
		stPis_CWOut.req_Close:=TRUE;
		
	END_IF
		
	IF NOT stPis_CWIn.st_Open THEN
		stPis_CWIn.req_Open:=TRUE;
	END_IF
	
ELSE
	IF NOT stPis_CWOut.st_Close THEN;
		stPis_CWOut.req_Close:=TRUE;
	END_IF
	
	IF NOT stPis_CWIn.st_Close THEN
		stPis_CWIn.req_Close:=TRUE;
	END_IF
END_IF
END_ACTION

PROPERTY cip_Pump_linked : BOOL
GET
cip_Pump_linked:=memo_CIP_Pump_linked;
END_GET
SET
memo_CIP_Pump_linked:=cip_Pump_linked;
END_SET
END_PROPERTY

METHOD m_Get_TriBlender_Clean : BOOL
VAR_INPUT
END_VAR
CASE eElementID OF
	E_Element_List.eTank_1,E_Element_List.eTank_2:;
		m_Get_TriBlender_Clean:=fbElement[E_Element_List.eTriBlender_Color].m_Get_State_Short()=E_Element_State_Short.eClean;
	E_Element_List.eTank_3,E_Element_List.eTank_4:;
		m_Get_TriBlender_Clean:=fbElement[E_Element_List.eTriBlender_Marinada].m_Get_State_Short()=E_Element_State_Short.eClean;
	
ELSE;
	m_Get_TriBlender_Clean:=FALSE;
END_CASE
END_METHOD

METHOD m_HMI : BOOL
VAR_INPUT
END_VAR
fbEvent_echo();
event_state_Update_sum:= TO_INT(eStatus) + TO_INT(stProdParam.eStatus) + TO_INT(eProcess);

IF event_state_Update_sum_last<>event_state_Update_sum THEN;
	event_state_Update_sum_last:=event_state_Update_sum;
	fbEvent_echo.event();
END_IF

event_state_Update:=fbEvent_echo.echo;
END_METHOD

METHOD m_Production_Run_Pump : BOOL
VAR_INPUT
END_VAR
CASE stProdParam.stRecipe.eFilling_Mode OF
	E_Filling_Mode.Line_Cyrculation,
	E_Filling_Mode.Bin_Cyrculation:;	
			IF TRUE
			AND trn_Tank_Color
			AND (refState_Long=E_Element_State_Long.eProduction
				OR (refState_Long=E_Element_State_Long.eExpired 
					AND refElement.eState_Long_Expiered =E_Element_State_Long.eProduction)
			AND fbTarget.m_CheckStatus(eReqStatus:=E_Tank_Target.eOpen)) 
			AND ((trn_Tank_A 
				AND fbLineSource.m_CheckStatus(eReqStatus:=E_Line_Source.eTank_A) 
				AND fbLineTarget.m_CheckStatus(eReqStatus:=E_Line_Target.eTank_A))
					OR
				(trn_Tank_B 
				AND fbLineSource.m_CheckStatus(eReqStatus:=E_Line_Source.eTank_B) 
				AND fbLineTarget.m_CheckStatus(eReqStatus:=E_Line_Target.eTank_B)))		
			AND fbInterConnection_ProL.bActive
			AND TRUE
			THEN;
				m_Production_Run_Pump:=TRUE;
			ELSE;
				m_Production_Run_Pump:=FALSE;
			END_IF	
	E_Filling_Mode.Bin:;
				m_Production_Run_Pump:=fbFilling.pumpFilling;
				
	E_Filling_Mode.Not_Selected:;
	
END_CASE
END_METHOD

METHOD m_Set_SFCFlags_Reference : BOOL
//Set reference to SFC flags

refSFC.SFCInit REF= SFCInit;
refSFC.SFCReset REF= SFCReset;
refSFC.SFCError REF= SFCError;
refSFC.SFCEnableLimit REF= SFCEnableLimit;
refSFC.SFCErrorStep REF= SFCErrorStep;
refSFC.SFCErrorPOU REF= SFCErrorPOU;
refSFC.SFCQuitError REF= SFCQuitError;
refSFC.SFCPause REF= SFCPause;
refSFC.SFCTrans REF= SFCTrans;
refSFC.SFCCurrentStep REF= SFCCurrentStep;
refSFC.SFCTip REF= SFCTip;
refSFC.SFCTipMode REF= SFCTipMode;

// Cycle handle for SFC
m_SFC_Handle();
END_METHOD

METHOD m_Stirrer : BOOL
VAR_INPUT
END_VAR
IF eStatus>=E_Element_State_Long.eWaterReady THEN;
	IF stProdParam.eStatus=E_Prod_Status.Active THEN;
		IF fbInterConnection_TriB.bActive THEN;
			m_Stirrer_run(param:=stProdParam.stRecipe.StirrerDissolving);
		ELSIF fbInterConnection_ProL.bActive THEN;
			IF memo_Production_Storage_Mode THEN;
				m_Stirrer_run(param:=stProdParam.stRecipe.StirrerStorage);
			ELSE;
				m_Stirrer_run(param:=stProdParam.stRecipe.StirrerProduction);
			END_IF	
		ELSE;		
			m_Stirrer_run(param:=stProdParam.stRecipe.StirrerStorage);//fb_Stirrer.m_Run(RPM:=1203);
		END_IF
	ELSE;
		fb_Stirrer.m_Run(RPM:=stProdParam.stRecipe.StirrerStorage.Speed);
	END_IF
ELSIF eStatus<E_Element_State_Long.eWaterReady
AND refElement.m_Get_InterConnection()=E_InterConnection.ConnToCIP THEN;
	// controled by CIP
	m_Stirrer_run_CIP();
ELSE;
	fb_Stirrer.m_Stop();
END_IF
END_METHOD

METHOD m_Stirrer_run : BOOL
VAR_INPUT
	param: ST_Prod_Param_Stirrer;
END_VAR

VAR
	time_on: TIME;
	time_off: TIME;
	time_cycle: TIME;
	
	dint_temp: DINT;
END_VAR
dint_temp:=param.tON*60000;
time_on:=TO_TIME(dint_temp);
dint_temp:=param.tOFF*60000;
time_off:=TO_TIME(dint_temp);
time_cycle:=time_on+time_off;
tonStirrer_time(PT:=time_cycle, IN:=NOT tonStirrer_time.Q);
IF tonStirrer_time.Q THEN;
	IF bStirrerDirectionPositive THEN;
		bStirrerDirectionPositive:=FALSE;
	ELSE;
		bStirrerDirectionPositive:=TRUE;
	END_IF
END_IF
CASE param.Mode OF 
	E_Stirrer_mode.continues:;
						fb_Stirrer.m_Run(RPM:=param.Speed);
	E_Stirrer_mode.cyclic:;
					IF tonStirrer_time.ET<time_on THEN;
						IF param.Flip_mode AND trn_Tank_Marinade THEN;
							IF bStirrerDirectionPositive THEN;
								fb_Stirrer.m_Run(RPM:=param.Speed);
							ELSE;
								fb_Stirrer.m_Run(RPM:=-param.Speed);
							END_IF							
						ELSE;
							fb_Stirrer.m_Run(RPM:=param.Speed);
						END_IF
						
					ELSE
						fb_Stirrer.m_Stop();
					END_IF
	E_Stirrer_mode.off:;
						fb_Stirrer.m_Stop();
END_CASE
END_METHOD

METHOD m_Stirrer_run_CIP : BOOL
VAR_INPUT
END_VAR
IF memo_CIP_Pump_linked
AND g_Pump.fbPump[E_Pump_List.P1001].bRun
THEN;
	fb_Stirrer.m_Run(RPM:=1204);
ELSE;
	fb_Stirrer.m_Stop();
END_IF
END_METHOD

METHOD mClearProduction : BOOL
VAR_INPUT
	state: E_Element_State_Long:=E_Element_State_Long.eOff;

END_VAR

VAR
	stRecipeEmpty: ST_Prod_Recipe;
END_VAR
stProdParam.eStatus:=E_Prod_Status.Not_Active;
stProdParam.stRecipe:=stRecipeEmpty;
eReq:=E_Request_List.eNone;

IF state<>E_Element_State_Long.eOff THEN;
	refState_Long:=state;
END_IF
END_METHOD

METHOD mGet_Recipe : BOOL
VAR_INPUT
	indexRecipe: INT;

END_VAR

VAR
	i: INT;
END_VAR
IF indexRecipe <0 OR indexRecipe > g_Prod.cMax_Prod_Recipe THEN;
	RETURN;
END_IF

CASE eElementID	OF 
	E_Element_List.eTank_1,E_Element_List.eTank_2:;
		stProdParam.stRecipe:=g_Prod.arrRecipeMarinade[indexRecipe];
	E_Element_List.eTank_3,E_Element_List.eTank_4:;
  		stProdParam.stRecipe:=g_Prod.arrRecipeColor[indexRecipe];
END_CASE

FOR i:=1 TO g_Prod.cMaxCompInProduct DO
	stProdParam.arrWeightIng[i]:=stProdParam.stRecipe.arr_Component[i].rWeightPercentage/100 * stProdParam.WeightOrder;
	stProdParam.stRecipe.arr_Component[i].rWeight:=stProdParam.stRecipe.arr_Component[i].rWeightPercentage/100 * stProdParam.WeightOrder;
END_FOR
END_METHOD

METHOD mTimeProductionDuration : TIME
VAR_INPUT
END_VAR
IF dtRealTime > stProdParam.prodDT 
AND stProdParam.eStatus=E_Prod_Status.Active
THEN;
	mTimeProductionDuration:=dtRealTime - stProdParam.prodDT;
ELSE;
	mTimeProductionDuration:=T#0S;
END_IF
END_METHOD

METHOD mTimeRemainToStart : TIME
VAR_INPUT
END_VAR
IF stProdParam.eStatus=E_Prod_Status.Activation_Pending_Shift THEN;
	stProdParam.eStatus:=E_Prod_Status.Activation_Pending;
	stProdParam.prodDT:=g_Prod.dtProdTimePicker+T#2h;
END_IF


IF stProdParam.eStatus=E_Prod_Status.Activation_Pending THEN;
	IF stProdParam.prodDT > dtRealTime THEN;
		mTimeRemainToStart:=stProdParam.prodDT - dtRealTime;
	ELSIF eStatus=E_Element_State_Long.eCIP_5_Done THEN;
		stProdParam.eStatus:=E_Prod_Status.Active;
		eReq:=E_Request_List.eWaterPrepare;
	END_IF
ELSE;
	mTimeRemainToStart:=T#0S;
END_IF
END_METHOD

PROPERTY pFilling_State : E_Filling_State
GET
pFilling_State:=eFilling_State;
END_GET
SET
eFilling_State:=pFilling_State;
END_SET
END_PROPERTY

TRANSITION trn_Tank_A:
trn_Tank_A:=(eElementID=E_Element_List.eTank_1 OR eElementID=E_Element_List.eTank_3);
END_TRANSITION

TRANSITION trn_Tank_B:
trn_Tank_B:=(eElementID=E_Element_List.eTank_2 OR eElementID=E_Element_List.eTank_4);
END_TRANSITION

TRANSITION trn_Tank_Color:
trn_Tank_Color:=(eElementID=E_Element_List.eTank_3 OR eElementID=E_Element_List.eTank_4);
END_TRANSITION

TRANSITION trn_Tank_Marinade:
trn_Tank_Marinade:=(eElementID=E_Element_List.eTank_1 OR eElementID=E_Element_List.eTank_2);
END_TRANSITION

END_FUNCTION_BLOCK

// ---- 00 Library/Sensors/FB_TankSensors.TcPOU
FUNCTION_BLOCK FB_TankSensors
VAR_IN_OUT
	stTankLevel	:	ST_Tank_Level	;
END_VAR
VAR_INPUT
	volume: REAL:=100; //litr
	//Level
	senHL				:	BOOL	;
	senLL				:	BOOL	;
	nSensorLvl_ID		: 	E_ASense_Name	;
	nSensorLvl_Raw		:	INT		;
	//Temperature
	nSensorTemp_ID		: 	E_ASense_Name	;
	nSensorTemp_Raw		:	INT		;
END_VAR
VAR_OUTPUT
	act_Volume			: REAL;
END_VAR
VAR
	stASensLvl			:	REFERENCE TO ST_AnalogSensor	;
	
	stASensTemp			:	REFERENCE TO ST_AnalogSensor	;
	
	Call_TankLevel			:	FB_AnalogSensor	;
	Call_TankTemp			:	FB_AnalogSensor	;
	tonEmpty: TON;
END_VAR

//Call_TankLevel(nSensorID:=nSensorLvl_ID, nRawSensor:=nSensorLvl_Raw );
//Call_TankTemp(nSensorID:=nSensorTemp_ID, nRawSensor:=nSensorTemp_Raw );
act_TankLvl();
act_Volume:=stTankLevel.rTankLevel;

ACTION act_TankLvl:
stASensLvl REF=g_AnalogSensor.stAnalogSensor[nSensorLvl_ID];

IF stTankLevel.bIn_LL_signal=FALSE AND stTankLevel.bIn_HL_signal=FALSE THEN
	tonEmpty.IN:=TRUE;
ELSE;
	tonEmpty.IN:=FALSE;
END_IF
IF stTankLevel.bIn_LL_signal=TRUE AND stTankLevel.bIn_HL_signal=FALSE THEN
	stTankLevel.e_state:=E_Tank_Level.eLL;
ELSIF stTankLevel.bIn_LL_signal=TRUE AND stTankLevel.bIn_HL_signal=TRUE THEN
	stTankLevel.e_state:=E_Tank_Level.eHL;
ELSIF stTankLevel.bIn_LL_signal=FALSE AND stTankLevel.bIn_HL_signal=TRUE THEN
	stTankLevel.e_state:=E_Tank_Level.eERROR;
END_IF

stTankLevel.rTankLevel:=stASensLvl.Value;
stTankLevel.rTankLevelPercentage:=stTankLevel.rTankLevel/volume*100;
stTankLevel.bIn_HL_signal:=senHL;
stTankLevel.bIn_LL_signal:=senLL;

tonEmpty(PT:=T#3S);
IF tonEmpty.Q THEN;
	stTankLevel.e_state:=E_Tank_Level.eEmpty;
END_IF
END_ACTION

METHOD get_stTankLevel : ST_Tank_Level
VAR_INPUT
END_VAR
VAR
	blank: ST_Tank_Level;
END_VAR
IF __ISVALIDREF(stTankLevel) THEN;
	get_stTankLevel:=stTankLevel;
ELSE;
	get_stTankLevel:=blank;
END_IF
END_METHOD

METHOD get_stTankLevel_OverFlow : BOOL
VAR_INPUT
END_VAR
VAR
	blank: ST_Tank_Level;
END_VAR
IF __ISVALIDREF(stTankLevel) THEN;
	IF stTankLevel.bIn_HL_signal 
	OR stTankLevel.rTankLevelPercentage>100
	OR (NOT MAIN.bTemp_Water_Overweight_check)
	THEN;
		get_stTankLevel_OverFlow:=TRUE;
	ELSE;
		get_stTankLevel_OverFlow:=FALSE;
	END_IF	
ELSE;
	get_stTankLevel_OverFlow:=FALSE;
END_IF
END_METHOD

END_FUNCTION_BLOCK

// ---- 00 Library/12 Analog Sensor/FB_AnalogSensor.TcPOU
FUNCTION_BLOCK FB_AnalogSensor
VAR_INPUT
	nSensorID	: 	E_ASense_Name	;
	nRawSensor	:	REAL				;
	arReset_AlrmWrn		:	ARRAY [0..3] OF BOOL		;//HH Alarm/LL Alarm/HH Warning/LL Warning
END_VAR
VAR_OUTPUT
	bLL_Alarm	:	BOOL	;
	bHH_Alarm	:	BOOL	;
	bLL_Warning	:	BOOL	;
	bHH_Warning	:	BOOL	;
END_VAR
VAR
	sName: STRING(12);

	stASens			:	REFERENCE TO ST_AnalogSensor	;
	state			: 	E_ASensor_State					;
	
	fbScaleFactor	: 	FB_ScaleFactor					;
	
	nTicks			:	INT:=0	;
	nI				:	INT		;
	
	bTestTemp		:	BOOL	;
	
	nTimeInCycles	:	INT:=100; //1 sec while cycletime is 10 ms
	nBufferSize_S	:	INT:=1	;//Buffer size in seconds
	nCycleTime_MS	:	INT:=10;//Cycle time in mili seconds
	
	
	//From Structure
	// Callibration 
	rawVal_Actual	: INT;//fb
	
	//MA
	arrRawVal_Actual	:	ARRAY [0..10000] OF INT	;//get out fb
	rTempRawVal			:	REAL	;//fb
	nRawSumm			:	DINT	;//fb
	
	bCopyRawTo_Min	: BOOL;//fb
	bCopyRawTo_Max	: BOOL;//fb
	
	//triggers
	arRS		:	ARRAY [0..3] OF RS		;//HH Alarm/LL Alarm/HH Warning/LL Warning
	
	ton_set_DATA: TON;
	rt_set_DATE: R_TRIG;
	fbScale: REFERENCE TO FB_ScaleFactor;
	fbMovingAverage: FB_MovingAverage;

	bSetFromTempCallibration: BOOL;
	bTypeTankConus: BOOL:=FALSE;
	rawTest: REAL;
END_VAR

nTimeInCycles:=TO_INT(nBufferSize_S*1000/nCycleTime_MS);
act_Get_Reference();
act_MA();
act_SetValues();
sName:=TO_STRING(nSensorID);
act_AlarmWarnings();

ACTION act_AlarmWarnings:
//arRS		:	ARRAY [0..3] OF RS		;//HH Alarm/LL Alarm/HH Warning/LL Warning
(*
arRS[0](
		SET:=(stASens.Value>= stASens.rHH_Alarm AND NOT bHH_Alarm) , 
		RESET1:=arReset_AlrmWrn[0] , Q1=>bHH_Alarm );
arRS[1](
		SET:=(stASens.Value<= stASens.rLL_Alarm AND NOT bLL_Alarm) , 
		RESET1:=arReset_AlrmWrn[1] , Q1=>bLL_Alarm );
arRS[2](
		SET:=(stASens.Value>= stASens.rHH_Warning AND stASens.Value<stASens.rHH_Alarm AND NOT bHH_Warning) , 
		RESET1:=arReset_AlrmWrn[2] , Q1=>bHH_Warning );
arRS[3](
		SET:=(stASens.Value<= stASens.rLL_Warning AND stASens.Value>stASens.rLL_Alarm AND NOT bLL_Warning) , 
		RESET1:=arReset_AlrmWrn[3] , Q1=>bLL_Warning );


*)		
bHH_Alarm:=stASens.Value>= stASens.rHH_Alarm;	
bLL_Alarm:=stASens.Value<= stASens.rLL_Alarm;	
bHH_Warning:=stASens.Value>= stASens.rHH_Warning AND stASens.Value<stASens.rHH_Alarm;	
bLL_Warning:=stASens.Value<= stASens.rLL_Warning AND stASens.Value>stASens.rLL_Alarm;
END_ACTION

ACTION act_Get_Reference:
stASens REF=g_AnalogSensor.stAnalogSensor[nSensorID];

stASens.ID:=TO_STRING(nSensorID);

//!!!!!!!!!!!!!!!!!!!!!!!!!!!!!!!!!!!!!!!!!!!!!!!!!!!!!!!!!!
//stASens.rawVal_Actual:=g_AnalogSensor.arAnalogSensorRawValue[nSensorID];
//stASens.rawVal_Actual:=nRawSensor;

//rTempRawVal:=rawTest;
CASE nSensorID OF 
	E_ASense_Name.LT3001,E_ASense_Name.LT3002,E_ASense_Name.LT4001,E_ASense_Name.LT4002:;
		bTypeTankConus:=TRUE;
ELSE;
		bTypeTankConus:=FALSE;
END_CASE
IF bTypeTankConus 
AND rTempRawVal<=stASens.rawVal_Min
THEN;
	stASens.Value:=mConus(rawValue:=rTempRawVal,baseIncriments:=stASens.rawVal_Min);
ELSE;
	fbScaleFactor(
		rVal:=rTempRawVal,//stASens.rawVal_Actual , 
		rInValHigh:=stASens.rawVal_Max , 
		rInValLow:=stASens.rawVal_Min , 
		rOutValHigh:=stASens.outVal_Max , 
		rOutValLow:=stASens.outVal_Min ,
		rOutOffset:=stASens.outOffset , 
		rValOut=>stASens.Value , 
		diValOut=>, 
		iValOut=> );	
END_IF

	
	
	
ton_set_DATA(PT:=T#20S, IN:=TRUE);
rt_set_DATE(CLK:=ton_set_DATA.Q);
IF rt_set_DATE.Q AND bSetFromTempCallibration THEN;
	set_Data(ID_reference:=nSensorID);
END_IF
END_ACTION

ACTION act_MA:
IF nTicks<nTimeInCycles THEN
	nTicks:=nTicks+1;
ELSIF nTicks>nTimeInCycles THEN
	nTicks:=nTimeInCycles;
END_IF

//moving ticks
nRawSumm:=0;
FOR nI:=nTimeInCycles TO 1 BY -1 DO
	arrRawVal_Actual[nI]:=arrRawVal_Actual[nI-1];
	//calculating summ
	nRawSumm:=nRawSumm+arrRawVal_Actual[nI];
END_FOR

arrRawVal_Actual[0]:=TO_INT(nRawSensor);
nRawSumm:=nRawSumm+arrRawVal_Actual[0];

rTempRawVal:=TO_REAL(nRawSumm/nTicks);


//fbMovingAverage(Value:=nRawSensor);
//rTempRawVal:=fbMovingAverage.Average;
END_ACTION

ACTION act_SetValues:
meth_SetRawValue(bSetValue:=bCopyRawTo_Max , nValToSet:=stASens.rawVal_Max , nRawValue:=rawVal_Actual );
meth_SetRawValue(bSetValue:=bCopyRawTo_Min , nValToSet:=stASens.rawVal_Min , nRawValue:=rawVal_Actual );
END_ACTION

METHOD mConus : REAL
VAR_INPUT
	rawValue: REAL;
	baseIncriments: REAL;
END_VAR



VAR
	hFactor: REAL;
	baseIncriment: REAL := 1050;
	h: REAL := 140;
	ConusConstant: REAL := 0.00000002165;
	pi: REAL:=3.1415926535;
	k: REAL:=3000000; // convert mm^3 to liters


	radius: REAL := 525;
	vConus: REAL;
END_VAR

VAR
	
END_VAR


//hFactor:=baseIncriment*h;

vConus:=pi*radius*radius*h/k;
IF baseIncriments=0 THEN;
	RETURN;
END_IF
ConusConstant:=vConus/(baseIncriments * baseIncriments * baseIncriments);
mConus:=ConusConstant*rawValue*rawValue*rawValue;
END_METHOD

METHOD INTERNAL meth_SetRawValue : BOOL
VAR_IN_OUT
	bSetValue	:	BOOL	;
	nValToSet	:	REAL	;
END_VAR
VAR_INPUT
	nRawValue	:	REAL		;
END_VAR
IF bSetValue THEN
	nValToSet:=nRawValue;
	bSetValue:=FALSE;
END_IF
END_METHOD

METHOD mSetAsConus : BOOL
VAR_INPUT
END_VAR
bTypeTankConus:=TRUE;
END_METHOD

METHOD set_Data : BOOL
VAR_INPUT
	ID_reference: E_ASense_Name;
END_VAR
fbScale REF= gIO.fbScaleFactor[ID_reference];
IF NOT __ISVALIDREF(fbScale) THEN;
	RETURN;
END_IF
	


stASens.rawVal_Max:=fbScale.rInValHigh;
stASens.rawVal_Min:=fbScale.rInValLow;
stASens.outVal_Max:=fbScale.rOutValHigh;
stASens.outVal_Min:=fbScale.rOutValLow;
stASens.outOffset:=fbScale.rOutOffset;
END_METHOD

END_FUNCTION_BLOCK

// ---- 00 Library/30 IO/FB_ScaleFactor.TcPOU
FUNCTION_BLOCK FB_ScaleFactor
VAR_INPUT
	rVal: REAL;
	rInValHigh: REAL;
	rInValLow: REAL;
	rOutValHigh: REAL;
	rOutValLow: REAL;
	rOutOffset: REAL:=0;
END_VAR

VAR
	rOfset: REAL;
	a: REAL;
	b: REAL;
END_VAR
VAR_OUTPUT
	rValOut: REAL;
	diValOut: DINT;
	iValOut: INT;
END_VAR

IF rInValHigh-rInValLow<>0 THEN;
	a:=(rOutValHigh-rOutValLow)/(rInValHigh-rInValLow);
ELSE;
	a:=0;
END_IF
b:=rOutValHigh-(a*rInValHigh);
rValOut:=(a*rVal+b)+rOutOffset;
diValOut:=TRUNC(rValOut);
iValOut:=DINT_TO_INT(diValOut);

END_FUNCTION_BLOCK

// ---- 00 Library/10 Utils/FB_MovingAverage.TcPOU
FUNCTION_BLOCK FB_MovingAverage
VAR_INPUT
	Value: REAL;
END_VAR
VAR_OUTPUT
	Average: REAL;

END_VAR
VAR
	arr: ARRAY[1..cMaxBufer] OF REAL;

	Sum: REAL;
	i: INT;
END_VAR
VAR CONSTANT
	cMaxBufer: INT:=500; // 10msec * 500 = 5 sec

END_VAR

Sum:=0;
FOR	i:=1 TO cMaxBufer DO
	Sum:=Sum+arr[i];
END_FOR


Average:=Sum/cMaxBufer;
FOR i:=cMaxBufer TO 2 BY-1 DO
	arr[i]:=arr[i-1];
END_FOR
arr[1]:=Value;

END_FUNCTION_BLOCK

// ---- 03 Project/11 Tank/FB_Filling.TcPOU
FUNCTION_BLOCK PUBLIC FB_Filling EXTENDS FB_SFC_Cycle IMPLEMENTS ITF_FB_SFC_Cycle
VAR_INPUT
	valFilling				: E_Pis_Name	;
	setWeight				: REAL:=200.0;	//kg
	actWeight				: REAL:=100.0;	//kg
	Tolerance				: REAL:=0.5;	//kg
	
END_VAR
VAR
	fbPis					: FB_Piston;	
	stPis_Filling			: REFERENCE TO ST_Piston;
	
	MinWeight	: REAL;
	MaxWeight	: REAL;
	
	reqTara		: BOOL;

END_VAR
VAR_IN_OUT
	eFill_State				: E_Filling_State;
END_VAR
VAR_OUTPUT
	eFill_State_HMI			: E_Filling_State;
	pumpFilling				: BOOL;
END_VAR

act_GetReference();

act_Oper();

MinWeight:=setWeight-Tolerance;
MaxWeight:=setWeight+Tolerance;
eFill_State_HMI:=eFill_State;

IF reqTara THEN;
	IF m_Tara() THEN;
		reqTara:=FALSE;
	ELSE;
		// tara command in process
	END_IF
END_IF

ACTION _aCheck_Condition_active:
// communication to weight


// check tara == weghit value <= 0.5 kg and >= -0.5 kg ==> 0 +- 0.5
bStepDone:=FALSE;
IF TRUE
//AND actWeight >= -0.5 AND actWeight <= 0.5 
AND actWeight < MinWeight 
AND eFill_State=E_Filling_State.eReady_ToFill
AND TRUE
THEN;
	bStepDone:=TRUE;
END_IF
END_ACTION

ACTION _aFilling_Process_active:
// check frow weight >= min value from recipe

pumpFilling:=m_FillingActive(); // Run autofiling process...
eFill_State:=E_Filling_State.eFilling_InProcess;

bStepDone:=FALSE;
IF actWeight >= MinWeight THEN;
	bStepDone:=TRUE;
END_IF
END_ACTION

ACTION _aFilling_Process_entry:
// open filling valve
fbPis.m_SetByRecipe(stPis:=stPis_Filling, 			req:=E_Piston_Recipe_State.Act);
// run pump
END_ACTION

ACTION _aFilling_Process_exit:
// close valve

// stop pump
END_ACTION

ACTION _aNo_Condition_active:
// print error
END_ACTION

ACTION _aReset_entry:
//close filing valve 
fbPis.m_SetByRecipe(stPis:=stPis_Filling, 			req:=E_Piston_Recipe_State.Release);

pumpFilling:=FALSE;
IF eFill_State=E_Filling_State.eFilling_InProcess THEN;
	eFill_State:=E_Filling_State.eReady_ToFill;
END_IF
bRun:=FALSE;
END_ACTION

ACTION act_GetReference:
m_Set_SFCFlags_Reference();

stPis_Filling				REF= g_Piston.stPis[valFilling];

(*
stPis_TankB				REF= g_Piston.stPis[valTankB];
stPis_TapWater			REF= g_Piston.stPis[valTapWater];
stPis_TapWater_else		REF= g_Piston.stPis[valTapWater_else];
stPis_TapWater_Drain	REF= g_Piston.stPis[valTapWater_Drain];
stPis_BlockWater		REF= g_Piston.stPis[valBlockWater];
stPis_WaterSource		REF= g_Piston.stPis[valWaterSource];
stPis_WaterSource_Drain	REF= g_Piston.stPis[valWaterSource_Drain];
stPis_Drain				REF= g_Piston.stPis[valDrain];
stPis_CIP				REF= g_Piston.stPis[valCIP];
stPis_CIP_Sel			REF= g_Piston.stPis[valCIP_Sel];
*)
END_ACTION

ACTION act_Oper:
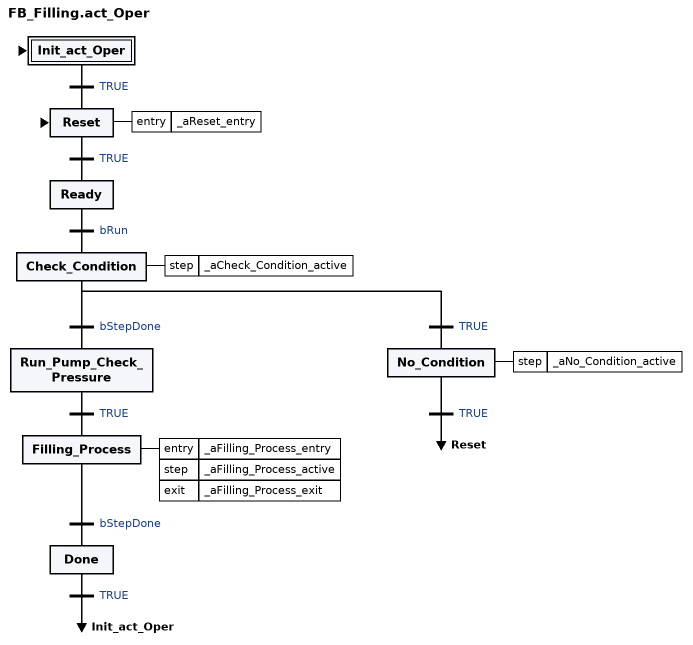
INITIAL_STEP Init_act_Oper:
END_STEP
TRANSITION FROM Init_act_Oper TO Reset
    := TRUE;
END_TRANSITION
STEP Reset:
    _aReset_entry(P1);  // entry action
END_STEP
TRANSITION FROM Reset TO Ready
    := TRUE;
END_TRANSITION
STEP Ready:
END_STEP
TRANSITION FROM Ready TO Check_Condition
    := bRun;
END_TRANSITION
STEP Check_Condition:
    _aCheck_Condition_active(N);  // step action
END_STEP
TRANSITION FROM Check_Condition TO Run_Pump_Check_Pressure
    := bStepDone;
END_TRANSITION
STEP Run_Pump_Check_Pressure:
END_STEP
TRANSITION FROM Run_Pump_Check_Pressure TO Filling_Process
    := TRUE;
END_TRANSITION
STEP Filling_Process:
    _aFilling_Process_entry(P1);  // entry action
    _aFilling_Process_active(N);  // step action
    _aFilling_Process_exit(P0);  // exit action
END_STEP
TRANSITION FROM Filling_Process TO Done
    := bStepDone;
END_TRANSITION
STEP Done:
END_STEP
TRANSITION FROM Done TO Init_act_Oper
    := TRUE;
END_TRANSITION
TRANSITION FROM Check_Condition TO No_Condition
    := TRUE;
END_TRANSITION
STEP No_Condition:  // min time T#2s
    _aNo_Condition_active(N);  // step action
END_STEP
TRANSITION FROM No_Condition TO Reset
    := TRUE;
END_TRANSITION
// branch label Branch0_act_Oper
END_ACTION

METHOD m_FillingActive : BOOL
VAR_INPUT
END_VAR

actWeight:=actWeight+0.1;
m_FillingActive:=TRUE;
END_METHOD

{warning 'add method implementation '}
METHOD m_Set_SFCFlags_Reference : BOOL
//Set reference to SFC flags

refSFC.SFCInit REF= SFCInit;
refSFC.SFCReset REF= SFCReset;
refSFC.SFCError REF= SFCError;
refSFC.SFCEnableLimit REF= SFCEnableLimit;
refSFC.SFCErrorStep REF= SFCErrorStep;
refSFC.SFCErrorPOU REF= SFCErrorPOU;
refSFC.SFCQuitError REF= SFCQuitError;
refSFC.SFCPause REF= SFCPause;
refSFC.SFCTrans REF= SFCTrans;
refSFC.SFCCurrentStep REF= SFCCurrentStep;
refSFC.SFCTip REF= SFCTip;
refSFC.SFCTipMode REF= SFCTipMode;

// Cycle handle for SFC
m_SFC_Handle();
END_METHOD

METHOD m_Tara : BOOL
VAR_INPUT
END_VAR
actWeight:=0.0;
m_Tara:=TRUE;
END_METHOD

END_FUNCTION_BLOCK

// ---- 03 Project/22 InterConnection/01 Tank/FB_Tank_Target.TcPOU
FUNCTION_BLOCK FB_Tank_Target EXTENDS FB_SFC_Cycle IMPLEMENTS ITF_FB_SFC_Cycle
VAR_INPUT
	//eElementID			: E_Element_List;
	valOutlet		: E_Pis_Name;
	valLine			: E_Pis_Name;
	valTriBlender	: E_Pis_Name;
	valDrain		: E_Pis_Name;	
	valCIP			: E_Pis_Name;	
END_VAR
VAR_OUTPUT
END_VAR
VAR
	//refElement		: REFERENCE TO FB_Element;
	//refState_Long		: REFERENCE TO E_Element_State_Long;
	eReq				: E_Tank_Target;
	eProcess			: E_Tank_Target;
	eStatus				: E_Tank_Target;
	
	fbPis				: FB_Piston;
	stPis_Outlet		: REFERENCE TO ST_Piston;
	stPis_Line			: REFERENCE TO ST_Piston;
	stPis_TriBlender	: REFERENCE TO ST_Piston;
	stPis_Drain			: REFERENCE TO ST_Piston;
	stPis_CIP			: REFERENCE TO ST_Piston;

	tonDrainTime: TON;
	rt_Req_Reset: R_TRIG;
	stTankLevel			:	ST_Tank_Level	;
END_VAR
VAR_IN_OUT


END_VAR

act_GetReference();

act_Oper();
IF NOT Init.x THEN;
	act_Status();
END_IF

tonDrainTime(PT:=T#1M, 
	IN:=(eStatus=E_Tank_Target.eDrain AND stTankLevel.e_state=E_Tank_Level.eEmpty)
			OR 
		eStatus=E_Tank_Target.eClose_DrainPipe);
IF tonDrainTime.Q 
AND eReq=E_Tank_Target.eNone
AND eProcess=E_Tank_Target.eNone
THEN;
	eReq:=E_Tank_Target.eClose;
END_IF

m_Request_Reset(memo:=rt_Req_Reset);//

ACTION _aCIP_active:
bStepDone:=FALSE;
IF TRUE 
AND eStatus=E_Tank_Target.eCIP
THEN;
	bStepDone:=TRUE;
END_IF
END_ACTION

ACTION _aCIP_entry:
fbPis.m_SetByRecipe(stPis:=stPis_Outlet, 		req:=E_Piston_Recipe_State.Act);
fbPis.m_SetByRecipe(stPis:=stPis_Line, 		req:=E_Piston_Recipe_State.Release);
fbPis.m_SetByRecipe(stPis:=stPis_TriBlender, 	req:=E_Piston_Recipe_State.Release);
fbPis.m_SetByRecipe(stPis:=stPis_Drain, 		req:=E_Piston_Recipe_State.Act);
fbPis.m_SetByRecipe(stPis:=stPis_CIP, 			req:=E_Piston_Recipe_State.Act);
END_ACTION

ACTION _aClose_active:
bStepDone:=FALSE;
IF TRUE 
AND eStatus=E_Tank_Target.eClose
THEN;
	bStepDone:=TRUE;
END_IF
END_ACTION

ACTION _aClose_entry:
fbPis.m_SetByRecipe(stPis:=stPis_Outlet, 		req:=E_Piston_Recipe_State.Release);
fbPis.m_SetByRecipe(stPis:=stPis_Line, 			req:=E_Piston_Recipe_State.Release);
fbPis.m_SetByRecipe(stPis:=stPis_TriBlender, 	req:=E_Piston_Recipe_State.Release);
fbPis.m_SetByRecipe(stPis:=stPis_Drain, 		req:=E_Piston_Recipe_State.Release);
fbPis.m_SetByRecipe(stPis:=stPis_CIP, 			req:=E_Piston_Recipe_State.Release);
END_ACTION

ACTION _aDone_entry:
eProcess:=E_Tank_Target.eNone;
eReq:=E_Tank_Target.eNone;
eStatus:=E_Tank_Target.eNone;
bRun:=FALSE;
bDone:=TRUE;
END_ACTION

ACTION _aDrain_active:
bStepDone:=FALSE;
IF TRUE 
AND eStatus=E_Tank_Target.eDrain
THEN;
	bStepDone:=TRUE;
END_IF
END_ACTION

ACTION _aDrain_entry:
fbPis.m_SetByRecipe(stPis:=stPis_Outlet, 		req:=E_Piston_Recipe_State.Act);
fbPis.m_SetByRecipe(stPis:=stPis_Line, 			req:=E_Piston_Recipe_State.Release);
fbPis.m_SetByRecipe(stPis:=stPis_TriBlender, 	req:=E_Piston_Recipe_State.Release);
fbPis.m_SetByRecipe(stPis:=stPis_Drain, 		req:=E_Piston_Recipe_State.Act);
fbPis.m_SetByRecipe(stPis:=stPis_CIP, 			req:=E_Piston_Recipe_State.Release);
END_ACTION

ACTION _aDrainPipe_active:
bStepDone:=FALSE;
IF TRUE 
AND eStatus=E_Tank_Target.eClose_DrainPipe
THEN;
	bStepDone:=TRUE;
END_IF
END_ACTION

ACTION _aDrainPipe_entry:
fbPis.m_SetByRecipe(stPis:=stPis_Outlet, 		req:=E_Piston_Recipe_State.Release);
fbPis.m_SetByRecipe(stPis:=stPis_Line, 			req:=E_Piston_Recipe_State.Release);
fbPis.m_SetByRecipe(stPis:=stPis_TriBlender, 	req:=E_Piston_Recipe_State.Release);
fbPis.m_SetByRecipe(stPis:=stPis_Drain, 		req:=E_Piston_Recipe_State.Act);
fbPis.m_SetByRecipe(stPis:=stPis_CIP, 			req:=E_Piston_Recipe_State.Release);
END_ACTION

ACTION _aInit_active:
SFCReset:=FALSE;
END_ACTION

ACTION _aInit_exit:
eProcess:=E_Tank_Target.eNone;
eReq:=E_Tank_Target.eNone;
END_ACTION

ACTION _aOpen_active:
bStepDone:=FALSE;
IF TRUE 
AND eStatus=E_Tank_Target.eOpen
THEN;
	bStepDone:=TRUE;
END_IF
END_ACTION

ACTION _aOpen_entry:
fbPis.m_SetByRecipe(stPis:=stPis_Outlet, req:=E_Piston_Recipe_State.Act);
//fbPis.m_SetByRecipe(stPis:=valLine, req:=E_Piston_Recipe_State.Release);
//fbPis.m_SetByRecipe(stPis:=valTriBlender, req:=E_Piston_Recipe_State.Release);
fbPis.m_SetByRecipe(stPis:=stPis_Drain, req:=E_Piston_Recipe_State.Release);
fbPis.m_SetByRecipe(stPis:=stPis_CIP, req:=E_Piston_Recipe_State.Release);
END_ACTION

ACTION _aReady_active:

eStatus:=E_Tank_Target.eNone;
CASE eReq OF
	E_Tank_Target.eClose:;
			IF TRUE THEN;
				eProcess:=E_Tank_Target.eClose;
			END_IF

	E_Tank_Target.eOpen:;
			IF TRUE THEN;
				eProcess:=E_Tank_Target.eOpen;
			END_IF	
			
	E_Tank_Target.eDrain:;
			IF TRUE THEN;
				eProcess:=E_Tank_Target.eDrain;
			END_IF
	
	E_Tank_Target.eClose_DrainPipe:;
			IF TRUE THEN;
				eProcess:=E_Tank_Target.eClose_DrainPipe;
			END_IF	
			
	E_Tank_Target.eCIP:;
			IF TRUE THEN;
				eProcess:=E_Tank_Target.eCIP;
			END_IF	

END_CASE
END_ACTION

ACTION _aReady_exit:
bRun:=TRUE;
bDone:=FALSE;
END_ACTION

ACTION act_GetReference:
m_Set_SFCFlags_Reference();
//refElement REF= fbElement[eElementID];
//refState_Long REF= fbElement[eElementID].eState_Long;

stPis_Outlet		REF= g_Piston.stPis[valOutlet];
stPis_Line			REF= g_Piston.stPis[valLine];
stPis_TriBlender	REF= g_Piston.stPis[valTriBlender];
stPis_Drain			REF= g_Piston.stPis[valDrain];
stPis_CIP			REF= g_Piston.stPis[valCIP];
END_ACTION

ACTION act_Oper:
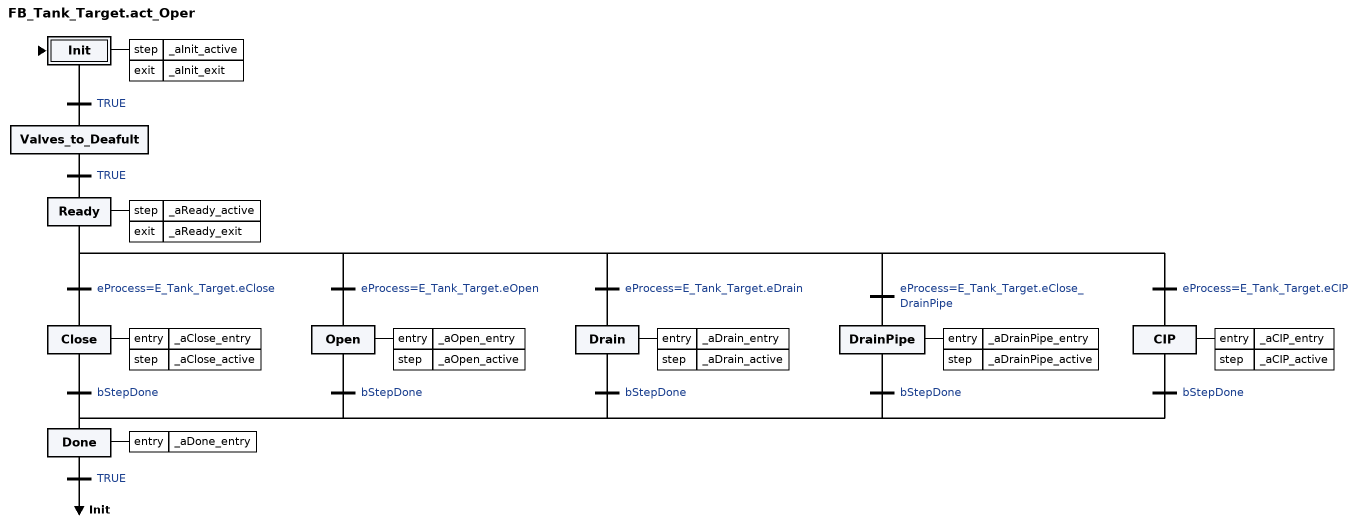
INITIAL_STEP Init:  // min time T#0.5s
    _aInit_active(N);  // step action
    _aInit_exit(P0);  // exit action
END_STEP
TRANSITION FROM Init TO Valves_to_Deafult
    := TRUE;
END_TRANSITION
STEP Valves_to_Deafult:
END_STEP
TRANSITION FROM Valves_to_Deafult TO Ready
    := TRUE;
END_TRANSITION
STEP Ready:
    _aReady_active(N);  // step action
    _aReady_exit(P0);  // exit action
END_STEP
TRANSITION FROM Ready TO Close
    := eProcess=E_Tank_Target.eClose;
END_TRANSITION
STEP Close:
    _aClose_entry(P1);  // entry action
    _aClose_active(N);  // step action
END_STEP
TRANSITION FROM Close TO Done
    := bStepDone;
END_TRANSITION
TRANSITION FROM Ready TO Open
    := eProcess=E_Tank_Target.eOpen;
END_TRANSITION
STEP Open:
    _aOpen_entry(P1);  // entry action
    _aOpen_active(N);  // step action
END_STEP
TRANSITION FROM Open TO Done
    := bStepDone;
END_TRANSITION
TRANSITION FROM Ready TO Drain
    := eProcess=E_Tank_Target.eDrain;
END_TRANSITION
STEP Drain:
    _aDrain_entry(P1);  // entry action
    _aDrain_active(N);  // step action
END_STEP
TRANSITION FROM Drain TO Done
    := bStepDone;
END_TRANSITION
TRANSITION FROM Ready TO DrainPipe
    := eProcess=E_Tank_Target.eClose_DrainPipe;
END_TRANSITION
STEP DrainPipe:
    _aDrainPipe_entry(P1);  // entry action
    _aDrainPipe_active(N);  // step action
END_STEP
TRANSITION FROM DrainPipe TO Done
    := bStepDone;
END_TRANSITION
TRANSITION FROM Ready TO CIP
    := eProcess=E_Tank_Target.eCIP;
END_TRANSITION
STEP CIP:
    _aCIP_entry(P1);  // entry action
    _aCIP_active(N);  // step action
END_STEP
TRANSITION FROM CIP TO Done
    := bStepDone;
END_TRANSITION
STEP Done:  // min time T#0.2s
    _aDone_entry(P1);  // entry action
END_STEP
TRANSITION FROM Done TO Init
    := TRUE;
END_TRANSITION
// branch label Branch0_act_Oper_Tank
END_ACTION

ACTION act_Status:


IF TRUE 
AND fbPis.m_CheckByRecipe(stPis:=stPis_Outlet, 		req:=E_Piston_Recipe_State.Release)
AND fbPis.m_CheckByRecipe(stPis:=stPis_Line, 		req:=E_Piston_Recipe_State.Release)
AND fbPis.m_CheckByRecipe(stPis:=stPis_TriBlender, 	req:=E_Piston_Recipe_State.Release)
AND fbPis.m_CheckByRecipe(stPis:=stPis_Drain, 		req:=E_Piston_Recipe_State.Release)
AND fbPis.m_CheckByRecipe(stPis:=stPis_CIP, 		req:=E_Piston_Recipe_State.Release)
THEN;
	eStatus:=E_Tank_Target.eClose;
	
ELSIF TRUE 
AND fbPis.m_CheckByRecipe(stPis:=stPis_Outlet, 		req:=E_Piston_Recipe_State.Act)
//AND fbPis.m_CheckByRecipe(stPis:=valLine, 		req:=E_Piston_Recipe_State.Release)
//AND fbPis.m_CheckByRecipe(stPis:=valTriBlender, 	req:=E_Piston_Recipe_State.Release)
AND fbPis.m_CheckByRecipe(stPis:=stPis_Drain, 		req:=E_Piston_Recipe_State.Release)
AND fbPis.m_CheckByRecipe(stPis:=stPis_CIP, 		req:=E_Piston_Recipe_State.Release)
THEN;
	eStatus:=E_Tank_Target.eOpen;
	
ELSIF TRUE 
AND fbPis.m_CheckByRecipe(stPis:=stPis_Outlet, 		req:=E_Piston_Recipe_State.Act)
AND fbPis.m_CheckByRecipe(stPis:=stPis_Line, 		req:=E_Piston_Recipe_State.Release)
AND fbPis.m_CheckByRecipe(stPis:=stPis_TriBlender, 	req:=E_Piston_Recipe_State.Release)
AND fbPis.m_CheckByRecipe(stPis:=stPis_Drain, 		req:=E_Piston_Recipe_State.Act)
AND fbPis.m_CheckByRecipe(stPis:=stPis_CIP, 		req:=E_Piston_Recipe_State.Release)
THEN;
	eStatus:=E_Tank_Target.eDrain;
	
ELSIF TRUE 
AND fbPis.m_CheckByRecipe(stPis:=stPis_Outlet, 		req:=E_Piston_Recipe_State.Release)
AND fbPis.m_CheckByRecipe(stPis:=stPis_Line, 		req:=E_Piston_Recipe_State.Release)
AND fbPis.m_CheckByRecipe(stPis:=stPis_TriBlender, 	req:=E_Piston_Recipe_State.Release)
AND fbPis.m_CheckByRecipe(stPis:=stPis_Drain, 		req:=E_Piston_Recipe_State.Act)
AND fbPis.m_CheckByRecipe(stPis:=stPis_CIP, 		req:=E_Piston_Recipe_State.Release)
THEN;
	eStatus:=E_Tank_Target.eClose_DrainPipe;
	
ELSIF TRUE 
AND fbPis.m_CheckByRecipe(stPis:=stPis_Outlet, 		req:=E_Piston_Recipe_State.Act)
AND fbPis.m_CheckByRecipe(stPis:=stPis_Line, 		req:=E_Piston_Recipe_State.Release)
AND fbPis.m_CheckByRecipe(stPis:=stPis_TriBlender, 	req:=E_Piston_Recipe_State.Release)
AND fbPis.m_CheckByRecipe(stPis:=stPis_Drain, 		req:=E_Piston_Recipe_State.Act)
AND fbPis.m_CheckByRecipe(stPis:=stPis_CIP, 		req:=E_Piston_Recipe_State.Act)
THEN;
	eStatus:=E_Tank_Target.eCIP;
	
ELSE;
	eStatus:=E_Tank_Target.eNone;
END_IF
END_ACTION

METHOD m_CheckStatus : BOOL
VAR_INPUT
	eReqStatus		: E_Tank_Target;
END_VAR
IF eStatus=eReqStatus 
AND eProcess=E_Tank_Target.eNone
AND eReq=E_Tank_Target.eNone
AND bReady
AND bDone
AND NOT bRun
THEN;
	m_CheckStatus:=TRUE;
END_IF
END_METHOD

METHOD m_Request_Reset : BOOL
VAR_IN_OUT
	memo: R_TRIG;
END_VAR
memo(CLK:=eReq=0);
IF TRUE 
AND memo.Q
THEN;
	SFCReset:=TRUE;
END_IF
END_METHOD

METHOD m_Run : BOOL
VAR_INPUT
	eReqProc			: E_Tank_Target;
END_VAR
IF eProcess=E_Tank_Target.eNone THEN;
	eProcess:=eReq:=eReqProc;
	bDone:=FALSE;
	m_Run:=TRUE;
END_IF
END_METHOD

METHOD m_Set_SFCFlags_Reference : BOOL
//Set reference to SFC flags

refSFC.SFCInit REF= SFCInit;
refSFC.SFCReset REF= SFCReset;
refSFC.SFCError REF= SFCError;
refSFC.SFCEnableLimit REF= SFCEnableLimit;
refSFC.SFCErrorStep REF= SFCErrorStep;
refSFC.SFCErrorPOU REF= SFCErrorPOU;
refSFC.SFCQuitError REF= SFCQuitError;
refSFC.SFCPause REF= SFCPause;
refSFC.SFCTrans REF= SFCTrans;
refSFC.SFCCurrentStep REF= SFCCurrentStep;
refSFC.SFCTip REF= SFCTip;
refSFC.SFCTipMode REF= SFCTipMode;

// Cycle handle for SFC
m_SFC_Handle();
END_METHOD

METHOD set_TankLevel : BOOL
VAR_INPUT
	set_stTankLevel			:	ST_Tank_Level	;
END_VAR
stTankLevel:=set_stTankLevel;
END_METHOD

END_FUNCTION_BLOCK

// ---- 03 Project/22 InterConnection/03 Line/FB_Line_Source.TcPOU
FUNCTION_BLOCK FB_Line_Source EXTENDS FB_SFC_Cycle IMPLEMENTS ITF_FB_SFC_Cycle
VAR_INPUT
	valTankA				:	E_Pis_Name	;
	valTankB				:	E_Pis_Name	;
	valTapWater				:	E_Pis_Name	;
	valTapWater_else		:	E_Pis_Name	;
	valTapWater_Drain		:	E_Pis_Name	;	
	valDrain				:	E_Pis_Name	;
	valCIP					:	E_Pis_Name	;
	valCIP_Sel				:	E_Pis_Name	;
	valBlockWater			:	E_Pis_Name	;	
	valWaterSource			:	E_Pis_Name	;
	valWaterSource_Drain	:	E_Pis_Name	;

END_VAR
VAR_OUTPUT
END_VAR
VAR
	eReq				: E_Line_Source;
	eProcess			: E_Line_Source;
	eStatus				: E_Line_Source;
	
	fbPis				: FB_Piston;
	
	stPis_TankA				: REFERENCE TO ST_Piston;
	stPis_TankB				: REFERENCE TO ST_Piston;
	stPis_TapWater			: REFERENCE TO ST_Piston;
	stPis_TapWater_else		: REFERENCE TO ST_Piston;
	stPis_TapWater_Drain	: REFERENCE TO ST_Piston;
	stPis_Drain				: REFERENCE TO ST_Piston;
	stPis_CIP				: REFERENCE TO ST_Piston;
	stPis_CIP_Sel			: REFERENCE TO ST_Piston;
	stPis_BlockWater		: REFERENCE TO ST_Piston;
	stPis_WaterSource		: REFERENCE TO ST_Piston;
	stPis_WaterSource_Drain	: REFERENCE TO ST_Piston;
	
	stPis_Outlet: ST_Piston;
	tonDrainTime: TON;
	ton_TapWaterNotInUse: TON;
	ton_TapWaterDrain_Timeout: TON;
	rt_Req_Reset: R_TRIG;
END_VAR

act_GetReference();

act_Oper();
//IF NOT Init.x THEN
	act_Status();
//END_IF

m_TapWaterNotInUse();

tonDrainTime(PT:=T#1M, IN:=eStatus=E_Line_Source.eDrain AND eReq=E_Line_Target.eNone);
IF tonDrainTime.Q 
AND eReq=E_Line_Source.eNone
AND eProcess=E_Line_Source.eNone
THEN;
	eReq:=E_Line_Source.eClose;
END_IF

m_Request_Reset(memo:=rt_Req_Reset);//

ACTION _aCIP_active:
bStepDone:=FALSE;
IF TRUE 
AND eStatus=E_Line_Source.eCIP
THEN;
	bStepDone:=TRUE;
END_IF
END_ACTION

ACTION _aCIP_entry:
fbPis.m_SetByRecipe(stPis:=stPis_TankA, 			req:=E_Piston_Recipe_State.Release);		
fbPis.m_SetByRecipe(stPis:=stPis_TankB, 			req:=E_Piston_Recipe_State.Release);
fbPis.m_SetByRecipe(stPis:=stPis_TapWater, 			req:=E_Piston_Recipe_State.Release);
fbPis.m_SetByRecipe(stPis:=stPis_TapWater_Drain, 	req:=E_Piston_Recipe_State.Release);
fbPis.m_SetByRecipe(stPis:=stPis_Drain, 			req:=E_Piston_Recipe_State.Act);
fbPis.m_SetByRecipe(stPis:=stPis_CIP, 				req:=E_Piston_Recipe_State.Act);
fbPis.m_SetByRecipe(stPis:=stPis_CIP_Sel,			req:=E_Piston_Recipe_State.Act);
fbPis.m_SetByRecipe(stPis:=stPis_BlockWater, 		req:=E_Piston_Recipe_State.Act);
fbPis.m_SetByRecipe(stPis:=stPis_WaterSource, 		req:=E_Piston_Recipe_State.Release);
fbPis.m_SetByRecipe(stPis:=stPis_WaterSource_Drain, req:=E_Piston_Recipe_State.Release);
END_ACTION

ACTION _aClose_active:
bStepDone:=FALSE;
IF TRUE 
AND eStatus=E_Line_Source.eClose
THEN;
	bStepDone:=TRUE;
END_IF
END_ACTION

ACTION _aClose_entry:
fbPis.m_SetByRecipe(stPis:=stPis_TankA, 			req:=E_Piston_Recipe_State.Release);		
fbPis.m_SetByRecipe(stPis:=stPis_TankB, 			req:=E_Piston_Recipe_State.Release);
fbPis.m_SetByRecipe(stPis:=stPis_TapWater, 			req:=E_Piston_Recipe_State.Release);
fbPis.m_SetByRecipe(stPis:=stPis_TapWater_Drain, 	req:=E_Piston_Recipe_State.Release);
fbPis.m_SetByRecipe(stPis:=stPis_Drain, 			req:=E_Piston_Recipe_State.Release);
fbPis.m_SetByRecipe(stPis:=stPis_CIP, 				req:=E_Piston_Recipe_State.Release);
fbPis.m_SetByRecipe(stPis:=stPis_CIP_Sel,			req:=E_Piston_Recipe_State.Release);
fbPis.m_SetByRecipe(stPis:=stPis_BlockWater, 		req:=E_Piston_Recipe_State.Release);
fbPis.m_SetByRecipe(stPis:=stPis_WaterSource, 		req:=E_Piston_Recipe_State.Release);
fbPis.m_SetByRecipe(stPis:=stPis_WaterSource_Drain, req:=E_Piston_Recipe_State.Release);
END_ACTION

ACTION _aDone_entry:
eProcess:=E_Line_Source.eNone;
eReq:=E_Line_Source.eNone;
bRun:=FALSE;
bDone:=TRUE;
END_ACTION

ACTION _aDrain_active:
bStepDone:=FALSE;
IF TRUE 
AND eStatus=E_Line_Source.eDrain
THEN;
	bStepDone:=TRUE;
END_IF
END_ACTION

ACTION _aDrain_entry:
fbPis.m_SetByRecipe(stPis:=stPis_TankA, 			req:=E_Piston_Recipe_State.Release);		
fbPis.m_SetByRecipe(stPis:=stPis_TankB, 			req:=E_Piston_Recipe_State.Release);
fbPis.m_SetByRecipe(stPis:=stPis_TapWater, 			req:=E_Piston_Recipe_State.Release);
fbPis.m_SetByRecipe(stPis:=stPis_TapWater_Drain, 	req:=E_Piston_Recipe_State.Release);
fbPis.m_SetByRecipe(stPis:=stPis_Drain, 			req:=E_Piston_Recipe_State.Act);
fbPis.m_SetByRecipe(stPis:=stPis_CIP, 				req:=E_Piston_Recipe_State.Release);
fbPis.m_SetByRecipe(stPis:=stPis_CIP_Sel,			req:=E_Piston_Recipe_State.Release);
fbPis.m_SetByRecipe(stPis:=stPis_BlockWater, 		req:=E_Piston_Recipe_State.Release);
fbPis.m_SetByRecipe(stPis:=stPis_WaterSource, 		req:=E_Piston_Recipe_State.Release);
fbPis.m_SetByRecipe(stPis:=stPis_WaterSource_Drain, req:=E_Piston_Recipe_State.Release);
END_ACTION

ACTION _aFill_Water_waiting_active:
bStepDone:=FALSE;
IF TRUE 
AND ton_TapWaterNotInUse.Q
THEN;
	bStepDone:=TRUE;
END_IF
END_ACTION

ACTION _aFillWater_active:
bStepDone:=FALSE;
IF TRUE 
AND eStatus=E_Line_Source.eFillWater
THEN;
	bStepDone:=TRUE;
END_IF
END_ACTION

ACTION _aFillWater_Drain_active:
;
END_ACTION

ACTION _aFillWater_Drain_entry:
fbPis.m_SetByRecipe(stPis:=stPis_TankA, 			req:=E_Piston_Recipe_State.Release);		
fbPis.m_SetByRecipe(stPis:=stPis_TankB, 			req:=E_Piston_Recipe_State.Release);
fbPis.m_SetByRecipe(stPis:=stPis_TapWater, 			req:=E_Piston_Recipe_State.Release);
fbPis.m_SetByRecipe(stPis:=stPis_TapWater_Drain, 	req:=E_Piston_Recipe_State.Release);
fbPis.m_SetByRecipe(stPis:=stPis_Drain, 			req:=E_Piston_Recipe_State.Release);
fbPis.m_SetByRecipe(stPis:=stPis_CIP, 				req:=E_Piston_Recipe_State.Release);
fbPis.m_SetByRecipe(stPis:=stPis_CIP_Sel,			req:=E_Piston_Recipe_State.Release);
fbPis.m_SetByRecipe(stPis:=stPis_BlockWater, 		req:=E_Piston_Recipe_State.Release);
fbPis.m_SetByRecipe(stPis:=stPis_WaterSource, 		req:=E_Piston_Recipe_State.Release);
fbPis.m_SetByRecipe(stPis:=stPis_WaterSource_Drain, req:=E_Piston_Recipe_State.Act);
END_ACTION

ACTION _aFillWater_entry:
fbPis.m_SetByRecipe(stPis:=stPis_TankA, 			req:=E_Piston_Recipe_State.Release);		
fbPis.m_SetByRecipe(stPis:=stPis_TankB, 			req:=E_Piston_Recipe_State.Release);
fbPis.m_SetByRecipe(stPis:=stPis_TapWater, 			req:=E_Piston_Recipe_State.Release);
fbPis.m_SetByRecipe(stPis:=stPis_TapWater_Drain, 	req:=E_Piston_Recipe_State.Release);
fbPis.m_SetByRecipe(stPis:=stPis_Drain, 			req:=E_Piston_Recipe_State.Release);
fbPis.m_SetByRecipe(stPis:=stPis_CIP, 				req:=E_Piston_Recipe_State.Release);
fbPis.m_SetByRecipe(stPis:=stPis_CIP_Sel,			req:=E_Piston_Recipe_State.Release);
fbPis.m_SetByRecipe(stPis:=stPis_BlockWater, 		req:=E_Piston_Recipe_State.Release);
fbPis.m_SetByRecipe(stPis:=stPis_WaterSource, 		req:=E_Piston_Recipe_State.Act);
fbPis.m_SetByRecipe(stPis:=stPis_WaterSource_Drain, req:=E_Piston_Recipe_State.Release);
END_ACTION

ACTION _aInit_active:
SFCReset:=FALSE;
END_ACTION

ACTION _aInit_exit:
eProcess:=E_Line_Source.eNone;
eReq:=E_Line_Source.eNone;
END_ACTION

ACTION _aReady_active:
CASE eReq OF
	E_Line_Source.eClose:;
			IF TRUE THEN;
				eProcess:=E_Line_Source.eClose;
			END_IF

	E_Line_Source.eTank_A:;
			IF TRUE THEN;
				eProcess:=E_Line_Source.eTank_A;
			END_IF	
			
	E_Line_Source.eTank_B:;
			IF TRUE THEN;
				eProcess:=E_Line_Source.eTank_B;
			END_IF	

	E_Line_Source.eTapWater:;
			IF TRUE THEN;
				eProcess:=E_Line_Source.eTapWater;
			END_IF	
			
	E_Line_Source.eFillWater:;
			IF TRUE THEN;
				eProcess:=E_Line_Source.eFillWater;
			END_IF	
			
	E_Line_Source.eCIP:;
			IF TRUE THEN;
				eProcess:=E_Line_Source.eCIP;
			END_IF	
			
	E_Line_Source.eDrain:;
			IF TRUE THEN;
				eProcess:=E_Line_Source.eDrain;
			END_IF			

END_CASE
END_ACTION

ACTION _aReady_exit:
bRun:=TRUE;
bDone:=FALSE;
END_ACTION

ACTION _aTank_A_active:
bStepDone:=FALSE;
IF TRUE 
AND eStatus=E_Line_Source.eTank_A
THEN;
	bStepDone:=TRUE;
END_IF
END_ACTION

ACTION _aTank_A_entry:
fbPis.m_SetByRecipe(stPis:=stPis_TankA, 			req:=E_Piston_Recipe_State.Act);		
fbPis.m_SetByRecipe(stPis:=stPis_TankB, 			req:=E_Piston_Recipe_State.Release);
fbPis.m_SetByRecipe(stPis:=stPis_TapWater, 			req:=E_Piston_Recipe_State.Release);
fbPis.m_SetByRecipe(stPis:=stPis_TapWater_Drain, 	req:=E_Piston_Recipe_State.Release);
fbPis.m_SetByRecipe(stPis:=stPis_Drain, 			req:=E_Piston_Recipe_State.Release);
fbPis.m_SetByRecipe(stPis:=stPis_CIP, 				req:=E_Piston_Recipe_State.Release);
fbPis.m_SetByRecipe(stPis:=stPis_CIP_Sel,			req:=E_Piston_Recipe_State.Release);
fbPis.m_SetByRecipe(stPis:=stPis_BlockWater, 		req:=E_Piston_Recipe_State.Act);
fbPis.m_SetByRecipe(stPis:=stPis_WaterSource, 		req:=E_Piston_Recipe_State.Release);
fbPis.m_SetByRecipe(stPis:=stPis_WaterSource_Drain, req:=E_Piston_Recipe_State.Release);
END_ACTION

ACTION _aTank_B_active:
bStepDone:=FALSE;
IF TRUE 
AND eStatus=E_Line_Source.eTank_B
THEN;
	bStepDone:=TRUE;
END_IF
END_ACTION

ACTION _aTank_B_entry:
fbPis.m_SetByRecipe(stPis:=stPis_TankA, 			req:=E_Piston_Recipe_State.Release);		
fbPis.m_SetByRecipe(stPis:=stPis_TankB, 			req:=E_Piston_Recipe_State.Act);
fbPis.m_SetByRecipe(stPis:=stPis_TapWater, 			req:=E_Piston_Recipe_State.Release);
fbPis.m_SetByRecipe(stPis:=stPis_TapWater_Drain, 	req:=E_Piston_Recipe_State.Release);
fbPis.m_SetByRecipe(stPis:=stPis_Drain, 			req:=E_Piston_Recipe_State.Release);
fbPis.m_SetByRecipe(stPis:=stPis_CIP, 				req:=E_Piston_Recipe_State.Release);
fbPis.m_SetByRecipe(stPis:=stPis_CIP_Sel,			req:=E_Piston_Recipe_State.Release);
fbPis.m_SetByRecipe(stPis:=stPis_BlockWater, 		req:=E_Piston_Recipe_State.Act);
fbPis.m_SetByRecipe(stPis:=stPis_WaterSource, 		req:=E_Piston_Recipe_State.Release);
fbPis.m_SetByRecipe(stPis:=stPis_WaterSource_Drain, 		req:=E_Piston_Recipe_State.Release);
END_ACTION

ACTION _aTap_Water_waiting_active:
bStepDone:=FALSE;
IF TRUE 
AND ton_TapWaterNotInUse.Q
THEN;
	bStepDone:=TRUE;
END_IF
END_ACTION

ACTION _aTapWater_active:
bStepDone:=FALSE;
IF TRUE 
AND eStatus=E_Line_Source.eTapWater
THEN;
	bStepDone:=TRUE;
END_IF
END_ACTION

ACTION _aTapWater_Drain_active:
//fbPis.m_SetByRecipe(stPis:=stPis_TapWater_Drain, 	req:=E_Piston_Recipe_State.Act);
END_ACTION

ACTION _aTapWater_Drain_entry:
fbPis.m_SetByRecipe(stPis:=stPis_TankA, 			req:=E_Piston_Recipe_State.Release);		
fbPis.m_SetByRecipe(stPis:=stPis_TankB, 			req:=E_Piston_Recipe_State.Release);
fbPis.m_SetByRecipe(stPis:=stPis_TapWater, 			req:=E_Piston_Recipe_State.Release);
fbPis.m_SetByRecipe(stPis:=stPis_TapWater_Drain, 	req:=E_Piston_Recipe_State.Act);
fbPis.m_SetByRecipe(stPis:=stPis_Drain, 			req:=E_Piston_Recipe_State.Release);
fbPis.m_SetByRecipe(stPis:=stPis_CIP, 				req:=E_Piston_Recipe_State.Release);
fbPis.m_SetByRecipe(stPis:=stPis_CIP_Sel,			req:=E_Piston_Recipe_State.Release);
fbPis.m_SetByRecipe(stPis:=stPis_BlockWater, 		req:=E_Piston_Recipe_State.Act);
fbPis.m_SetByRecipe(stPis:=stPis_WaterSource, 		req:=E_Piston_Recipe_State.Release);
fbPis.m_SetByRecipe(stPis:=stPis_WaterSource_Drain, req:=E_Piston_Recipe_State.Release);
END_ACTION

ACTION _aTapWater_entry:
fbPis.m_SetByRecipe(stPis:=stPis_TankA, 			req:=E_Piston_Recipe_State.Release);		
fbPis.m_SetByRecipe(stPis:=stPis_TankB, 			req:=E_Piston_Recipe_State.Release);
fbPis.m_SetByRecipe(stPis:=stPis_TapWater, 			req:=E_Piston_Recipe_State.Act);
fbPis.m_SetByRecipe(stPis:=stPis_TapWater_Drain, 	req:=E_Piston_Recipe_State.Release);
fbPis.m_SetByRecipe(stPis:=stPis_Drain, 			req:=E_Piston_Recipe_State.Release);
fbPis.m_SetByRecipe(stPis:=stPis_CIP, 				req:=E_Piston_Recipe_State.Release);
fbPis.m_SetByRecipe(stPis:=stPis_CIP_Sel,			req:=E_Piston_Recipe_State.Release);
fbPis.m_SetByRecipe(stPis:=stPis_BlockWater, 		req:=E_Piston_Recipe_State.Act);
fbPis.m_SetByRecipe(stPis:=stPis_WaterSource, 		req:=E_Piston_Recipe_State.Release);
fbPis.m_SetByRecipe(stPis:=stPis_WaterSource_Drain, req:=E_Piston_Recipe_State.Release);
END_ACTION

ACTION act_GetReference:
m_Set_SFCFlags_Reference();

stPis_TankA				REF= g_Piston.stPis[valTankA];
stPis_TankB				REF= g_Piston.stPis[valTankB];
stPis_TapWater			REF= g_Piston.stPis[valTapWater];
stPis_TapWater_else		REF= g_Piston.stPis[valTapWater_else];
stPis_TapWater_Drain	REF= g_Piston.stPis[valTapWater_Drain];
stPis_BlockWater		REF= g_Piston.stPis[valBlockWater];
stPis_WaterSource		REF= g_Piston.stPis[valWaterSource];
stPis_WaterSource_Drain	REF= g_Piston.stPis[valWaterSource_Drain];
stPis_Drain				REF= g_Piston.stPis[valDrain];
stPis_CIP				REF= g_Piston.stPis[valCIP];
stPis_CIP_Sel			REF= g_Piston.stPis[valCIP_Sel];
END_ACTION

ACTION act_Oper:
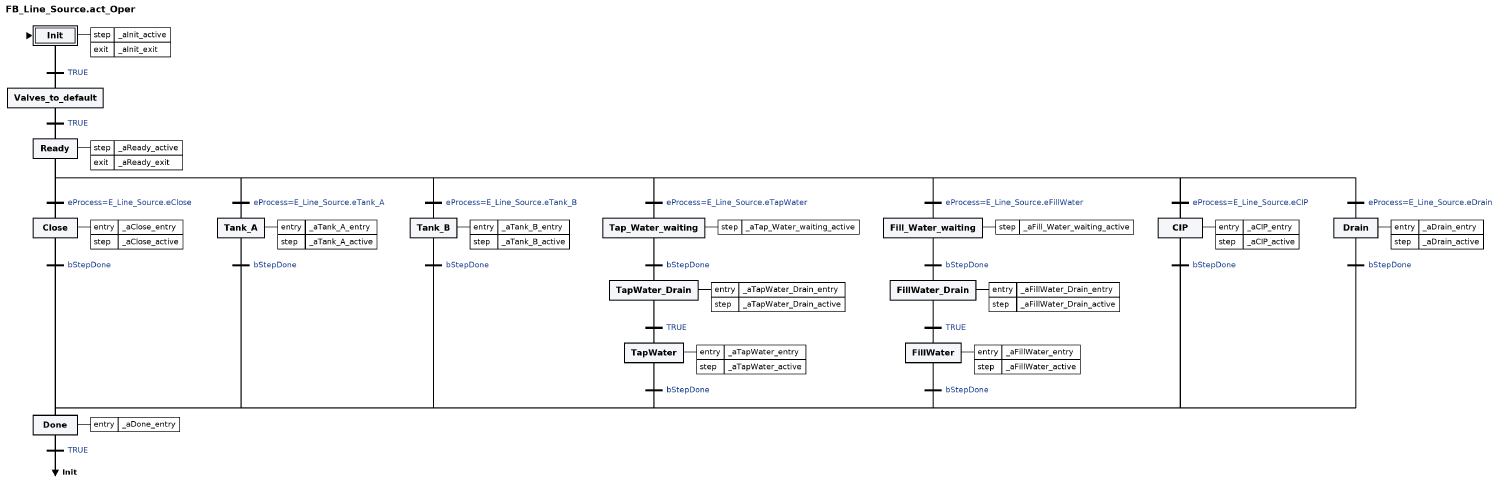
INITIAL_STEP Init:
    _aInit_active(N);  // step action
    _aInit_exit(P0);  // exit action
END_STEP
TRANSITION FROM Init TO Valves_to_default
    := TRUE;
END_TRANSITION
STEP Valves_to_default:
END_STEP
TRANSITION FROM Valves_to_default TO Ready
    := TRUE;
END_TRANSITION
STEP Ready:
    _aReady_active(N);  // step action
    _aReady_exit(P0);  // exit action
END_STEP
TRANSITION FROM Ready TO Close
    := eProcess=E_Line_Source.eClose;
END_TRANSITION
STEP Close:
    _aClose_entry(P1);  // entry action
    _aClose_active(N);  // step action
END_STEP
TRANSITION FROM Close TO Done
    := bStepDone;
END_TRANSITION
TRANSITION FROM Ready TO Tank_A
    := eProcess=E_Line_Source.eTank_A;
END_TRANSITION
STEP Tank_A:
    _aTank_A_entry(P1);  // entry action
    _aTank_A_active(N);  // step action
END_STEP
TRANSITION FROM Tank_A TO Done
    := bStepDone;
END_TRANSITION
TRANSITION FROM Ready TO Tank_B
    := eProcess=E_Line_Source.eTank_B;
END_TRANSITION
STEP Tank_B:
    _aTank_B_entry(P1);  // entry action
    _aTank_B_active(N);  // step action
END_STEP
TRANSITION FROM Tank_B TO Done
    := bStepDone;
END_TRANSITION
TRANSITION FROM Ready TO Tap_Water_waiting
    := eProcess=E_Line_Source.eTapWater;
END_TRANSITION
STEP Tap_Water_waiting:
    _aTap_Water_waiting_active(N);  // step action
END_STEP
TRANSITION FROM Tap_Water_waiting TO TapWater_Drain
    := bStepDone;
END_TRANSITION
STEP TapWater_Drain:  // min time T#10s
    _aTapWater_Drain_entry(P1);  // entry action
    _aTapWater_Drain_active(N);  // step action
END_STEP
TRANSITION FROM TapWater_Drain TO TapWater
    := TRUE;
END_TRANSITION
STEP TapWater:
    _aTapWater_entry(P1);  // entry action
    _aTapWater_active(N);  // step action
END_STEP
TRANSITION FROM TapWater TO Done
    := bStepDone;
END_TRANSITION
TRANSITION FROM Ready TO Fill_Water_waiting
    := eProcess=E_Line_Source.eFillWater;
END_TRANSITION
STEP Fill_Water_waiting:
    _aFill_Water_waiting_active(N);  // step action
END_STEP
TRANSITION FROM Fill_Water_waiting TO FillWater_Drain
    := bStepDone;
END_TRANSITION
STEP FillWater_Drain:  // min time T#10s
    _aFillWater_Drain_entry(P1);  // entry action
    _aFillWater_Drain_active(N);  // step action
END_STEP
TRANSITION FROM FillWater_Drain TO FillWater
    := TRUE;
END_TRANSITION
STEP FillWater:
    _aFillWater_entry(P1);  // entry action
    _aFillWater_active(N);  // step action
END_STEP
TRANSITION FROM FillWater TO Done
    := bStepDone;
END_TRANSITION
TRANSITION FROM Ready TO CIP
    := eProcess=E_Line_Source.eCIP;
END_TRANSITION
STEP CIP:
    _aCIP_entry(P1);  // entry action
    _aCIP_active(N);  // step action
END_STEP
TRANSITION FROM CIP TO Done
    := bStepDone;
END_TRANSITION
TRANSITION FROM Ready TO Drain
    := eProcess=E_Line_Source.eDrain;
END_TRANSITION
STEP Drain:
    _aDrain_entry(P1);  // entry action
    _aDrain_active(N);  // step action
END_STEP
TRANSITION FROM Drain TO Done
    := bStepDone;
END_TRANSITION
STEP Done:
    _aDone_entry(P1);  // entry action
END_STEP
TRANSITION FROM Done TO Init
    := TRUE;
END_TRANSITION
// branch label Branch0_act_Oper
END_ACTION

ACTION act_Status:
IF TRUE 
AND fbPis.m_CheckByRecipe(stPis:=stPis_TankA, 			req:=E_Piston_Recipe_State.Release)		
AND fbPis.m_CheckByRecipe(stPis:=stPis_TankB, 			req:=E_Piston_Recipe_State.Release)
AND fbPis.m_CheckByRecipe(stPis:=stPis_TapWater, 		req:=E_Piston_Recipe_State.Release)
AND fbPis.m_CheckByRecipe(stPis:=stPis_TapWater_Drain, 	req:=E_Piston_Recipe_State.Release)
AND fbPis.m_CheckByRecipe(stPis:=stPis_Drain, 			req:=E_Piston_Recipe_State.Release)
AND fbPis.m_CheckByRecipe(stPis:=stPis_CIP, 			req:=E_Piston_Recipe_State.Release)
AND fbPis.m_CheckByRecipe(stPis:=stPis_CIP_Sel,			req:=E_Piston_Recipe_State.Release)
AND fbPis.m_CheckByRecipe(stPis:=stPis_BlockWater, 		req:=E_Piston_Recipe_State.Release)
AND fbPis.m_CheckByRecipe(stPis:=stPis_WaterSource, 	req:=E_Piston_Recipe_State.Release)
AND fbPis.m_CheckByRecipe(stPis:=stPis_WaterSource_Drain,req:=E_Piston_Recipe_State.Release)
THEN;
	eStatus:=E_Line_Source.eClose;
ELSIF TRUE 
AND fbPis.m_CheckByRecipe(stPis:=stPis_TankA, 			req:=E_Piston_Recipe_State.Act)		
AND fbPis.m_CheckByRecipe(stPis:=stPis_TankB, 			req:=E_Piston_Recipe_State.Release)
AND fbPis.m_CheckByRecipe(stPis:=stPis_TapWater, 		req:=E_Piston_Recipe_State.Release)
AND fbPis.m_CheckByRecipe(stPis:=stPis_TapWater_Drain, 	req:=E_Piston_Recipe_State.Release)
AND fbPis.m_CheckByRecipe(stPis:=stPis_Drain, 			req:=E_Piston_Recipe_State.Release)
AND fbPis.m_CheckByRecipe(stPis:=stPis_CIP, 			req:=E_Piston_Recipe_State.Release)
AND fbPis.m_CheckByRecipe(stPis:=stPis_CIP_Sel,			req:=E_Piston_Recipe_State.Release)
AND fbPis.m_CheckByRecipe(stPis:=stPis_BlockWater, 		req:=E_Piston_Recipe_State.Act)
AND fbPis.m_CheckByRecipe(stPis:=stPis_WaterSource, 	req:=E_Piston_Recipe_State.Release)
AND fbPis.m_CheckByRecipe(stPis:=stPis_WaterSource_Drain,req:=E_Piston_Recipe_State.Release)
THEN;
	eStatus:=E_Line_Source.eTank_A;
ELSIF TRUE 
AND fbPis.m_CheckByRecipe(stPis:=stPis_TankA, 			req:=E_Piston_Recipe_State.Release)		
AND fbPis.m_CheckByRecipe(stPis:=stPis_TankB, 			req:=E_Piston_Recipe_State.Act)
AND fbPis.m_CheckByRecipe(stPis:=stPis_TapWater, 		req:=E_Piston_Recipe_State.Release)
AND fbPis.m_CheckByRecipe(stPis:=stPis_TapWater_Drain, 	req:=E_Piston_Recipe_State.Release)
AND fbPis.m_CheckByRecipe(stPis:=stPis_Drain, 			req:=E_Piston_Recipe_State.Release)
AND fbPis.m_CheckByRecipe(stPis:=stPis_CIP, 			req:=E_Piston_Recipe_State.Release)
AND fbPis.m_CheckByRecipe(stPis:=stPis_CIP_Sel,			req:=E_Piston_Recipe_State.Release)
AND fbPis.m_CheckByRecipe(stPis:=stPis_BlockWater, 		req:=E_Piston_Recipe_State.Act)
AND fbPis.m_CheckByRecipe(stPis:=stPis_WaterSource, 	req:=E_Piston_Recipe_State.Release)
AND fbPis.m_CheckByRecipe(stPis:=stPis_WaterSource_Drain,req:=E_Piston_Recipe_State.Release)
THEN;
	eStatus:=E_Line_Source.eTank_B;
ELSIF TRUE 
AND fbPis.m_CheckByRecipe(stPis:=stPis_TankA, 			req:=E_Piston_Recipe_State.Release)		
AND fbPis.m_CheckByRecipe(stPis:=stPis_TankB, 			req:=E_Piston_Recipe_State.Release)
AND fbPis.m_CheckByRecipe(stPis:=stPis_TapWater, 		req:=E_Piston_Recipe_State.Act)
AND fbPis.m_CheckByRecipe(stPis:=stPis_TapWater_Drain, 	req:=E_Piston_Recipe_State.Release)
AND fbPis.m_CheckByRecipe(stPis:=stPis_TapWater_else, 	req:=E_Piston_Recipe_State.Release)
AND fbPis.m_CheckByRecipe(stPis:=stPis_Drain, 			req:=E_Piston_Recipe_State.Release)
AND fbPis.m_CheckByRecipe(stPis:=stPis_CIP, 			req:=E_Piston_Recipe_State.Release)
AND fbPis.m_CheckByRecipe(stPis:=stPis_CIP_Sel,			req:=E_Piston_Recipe_State.Release)
AND fbPis.m_CheckByRecipe(stPis:=stPis_BlockWater, 		req:=E_Piston_Recipe_State.Act)
AND fbPis.m_CheckByRecipe(stPis:=stPis_WaterSource, 	req:=E_Piston_Recipe_State.Release)
AND fbPis.m_CheckByRecipe(stPis:=stPis_WaterSource_Drain,req:=E_Piston_Recipe_State.Release)
THEN;
	eStatus:=E_Line_Source.eTapWater;
ELSIF TRUE 
AND fbPis.m_CheckByRecipe(stPis:=stPis_TankA, 			req:=E_Piston_Recipe_State.Release)		
AND fbPis.m_CheckByRecipe(stPis:=stPis_TankB, 			req:=E_Piston_Recipe_State.Release)
AND fbPis.m_CheckByRecipe(stPis:=stPis_TapWater, 		req:=E_Piston_Recipe_State.Release)
AND fbPis.m_CheckByRecipe(stPis:=stPis_TapWater_Drain, 	req:=E_Piston_Recipe_State.Release)
AND fbPis.m_CheckByRecipe(stPis:=stPis_Drain, 			req:=E_Piston_Recipe_State.Release)
AND fbPis.m_CheckByRecipe(stPis:=stPis_CIP, 			req:=E_Piston_Recipe_State.Release)
AND fbPis.m_CheckByRecipe(stPis:=stPis_CIP_Sel,			req:=E_Piston_Recipe_State.Release)
AND fbPis.m_CheckByRecipe(stPis:=stPis_BlockWater, 		req:=E_Piston_Recipe_State.Release)
AND fbPis.m_CheckByRecipe(stPis:=stPis_WaterSource, 	req:=E_Piston_Recipe_State.Act)
AND fbPis.m_CheckByRecipe(stPis:=stPis_WaterSource_Drain,req:=E_Piston_Recipe_State.Release)
THEN;
	eStatus:=E_Line_Source.eFillWater;
ELSIF TRUE 
AND fbPis.m_CheckByRecipe(stPis:=stPis_TankA, 			req:=E_Piston_Recipe_State.Release)		
AND fbPis.m_CheckByRecipe(stPis:=stPis_TankB, 			req:=E_Piston_Recipe_State.Release)
AND fbPis.m_CheckByRecipe(stPis:=stPis_TapWater, 		req:=E_Piston_Recipe_State.Release)
AND fbPis.m_CheckByRecipe(stPis:=stPis_TapWater_Drain, 	req:=E_Piston_Recipe_State.Release)
AND fbPis.m_CheckByRecipe(stPis:=stPis_Drain, 			req:=E_Piston_Recipe_State.Act)
AND fbPis.m_CheckByRecipe(stPis:=stPis_CIP, 			req:=E_Piston_Recipe_State.Act)
AND fbPis.m_CheckByRecipe(stPis:=stPis_CIP_Sel,			req:=E_Piston_Recipe_State.Act)
AND fbPis.m_CheckByRecipe(stPis:=stPis_BlockWater, 		req:=E_Piston_Recipe_State.Act)
AND fbPis.m_CheckByRecipe(stPis:=stPis_WaterSource, 	req:=E_Piston_Recipe_State.Release)
AND fbPis.m_CheckByRecipe(stPis:=stPis_WaterSource_Drain,req:=E_Piston_Recipe_State.Release)
THEN;
	eStatus:=E_Line_Source.eCIP;
ELSIF TRUE 
AND fbPis.m_CheckByRecipe(stPis:=stPis_TankA, 			req:=E_Piston_Recipe_State.Release)		
AND fbPis.m_CheckByRecipe(stPis:=stPis_TankB, 			req:=E_Piston_Recipe_State.Release)
AND fbPis.m_CheckByRecipe(stPis:=stPis_TapWater, 		req:=E_Piston_Recipe_State.Release)
AND fbPis.m_CheckByRecipe(stPis:=stPis_TapWater_Drain, 	req:=E_Piston_Recipe_State.Release)
AND fbPis.m_CheckByRecipe(stPis:=stPis_Drain, 			req:=E_Piston_Recipe_State.Act)
AND fbPis.m_CheckByRecipe(stPis:=stPis_CIP, 			req:=E_Piston_Recipe_State.Release)
AND fbPis.m_CheckByRecipe(stPis:=stPis_CIP_Sel,			req:=E_Piston_Recipe_State.Release)
AND fbPis.m_CheckByRecipe(stPis:=stPis_BlockWater, 		req:=E_Piston_Recipe_State.Release)
AND fbPis.m_CheckByRecipe(stPis:=stPis_WaterSource, 	req:=E_Piston_Recipe_State.Release)
AND fbPis.m_CheckByRecipe(stPis:=stPis_WaterSource_Drain,req:=E_Piston_Recipe_State.Release)
THEN;
	eStatus:=E_Line_Source.eDrain;
ELSE;
	eStatus:=E_Line_Source.eNone;
END_IF
END_ACTION

METHOD m_CheckStatus : BOOL
VAR_INPUT
	eReqStatus		: E_Line_Source;
END_VAR
IF eStatus=eReqStatus 
AND eProcess=E_Line_Source.eNone
AND eReq=E_Line_Source.eNone
AND bReady
AND bDone
AND NOT bRun
THEN;
	m_CheckStatus:=TRUE;
END_IF
END_METHOD

METHOD m_Request_Reset : BOOL
VAR_IN_OUT
	memo: R_TRIG;
END_VAR
memo(CLK:=eReq=0);
IF TRUE 
AND memo.Q
THEN;
	SFCReset:=TRUE;
END_IF
END_METHOD

METHOD m_Run : BOOL
VAR_INPUT
	eReqProc			: E_Line_Source;
END_VAR
IF eProcess=E_Line_Source.eNone THEN;
	eProcess:=eReq:=eReqProc;
	bDone:=FALSE;
	m_Run:=TRUE;
END_IF
END_METHOD

METHOD m_Set_SFCFlags_Reference : BOOL
//Set reference to SFC flags

refSFC.SFCInit REF= SFCInit;
refSFC.SFCReset REF= SFCReset;
refSFC.SFCError REF= SFCError;
refSFC.SFCEnableLimit REF= SFCEnableLimit;
refSFC.SFCErrorStep REF= SFCErrorStep;
refSFC.SFCErrorPOU REF= SFCErrorPOU;
refSFC.SFCQuitError REF= SFCQuitError;
refSFC.SFCPause REF= SFCPause;
refSFC.SFCTrans REF= SFCTrans;
refSFC.SFCCurrentStep REF= SFCCurrentStep;
refSFC.SFCTip REF= SFCTip;
refSFC.SFCTipMode REF= SFCTipMode;

// Cycle handle for SFC
m_SFC_Handle();
END_METHOD

METHOD m_TapWaterNotInUse : BOOL
VAR_INPUT
END_VAR
IF TRUE 
AND fbPis.m_CheckByRecipe(stPis:=stPis_TapWater, 			req:=E_Piston_Recipe_State.Release)		
AND fbPis.m_CheckByRecipe(stPis:=stPis_TapWater_Drain, 		req:=E_Piston_Recipe_State.Release)
AND fbPis.m_CheckByRecipe(stPis:=stPis_TapWater_else, 		req:=E_Piston_Recipe_State.Release)
AND fbPis.m_CheckByRecipe(stPis:=stPis_WaterSource, 		req:=E_Piston_Recipe_State.Release)
AND fbPis.m_CheckByRecipe(stPis:=stPis_WaterSource_Drain, 	req:=E_Piston_Recipe_State.Release)
THEN;
	ton_TapWaterNotInUse(IN:=TRUE);
ELSE;
	ton_TapWaterNotInUse(IN:=FALSE);
END_IF

ton_TapWaterNotInUse(PT:=T#3S);


//Tap Water Drain Timeout
ton_TapWaterDrain_Timeout(PT:=T#10S);
IF fbPis.m_CheckByRecipe(stPis:=stPis_TapWater_Drain, 	req:=E_Piston_Recipe_State.Act) THEN;
	ton_TapWaterDrain_Timeout.IN:=TRUE;
ELSE;
	ton_TapWaterDrain_Timeout.IN:=FALSE;
END_IF
IF ton_TapWaterDrain_Timeout.Q THEN;
	fbPis.m_SetByRecipe(stPis:=stPis_TapWater_Drain, 	req:=E_Piston_Recipe_State.Release);
END_IF
END_METHOD

END_FUNCTION_BLOCK

// ---- 03 Project/22 InterConnection/03 Line/FB_Line_Target.TcPOU
FUNCTION_BLOCK FB_Line_Target EXTENDS FB_SFC_Cycle IMPLEMENTS ITF_FB_SFC_Cycle
VAR_INPUT
	valTankA				:	E_Pis_Name	;
	valTankB				:	E_Pis_Name	;
	valTankA_Pipe			:	E_Pis_Name	;
	valTankB_Pipe			:	E_Pis_Name	;
	valDrain				:	E_Pis_Name	;
	valCIP					:	E_Pis_Name	;
END_VAR
VAR_OUTPUT
END_VAR
VAR
	eReq				: E_Line_Target;
	eProcess			: E_Line_Target;
	eStatus				: E_Line_Target;
	
	fbPis				: FB_Piston;
	
	stPis_TankA				: REFERENCE TO ST_Piston;
	stPis_TankB				: REFERENCE TO ST_Piston;
	stPis_TankA_Pipe		: REFERENCE TO ST_Piston;
	stPis_TankB_Pipe		: REFERENCE TO ST_Piston;
	stPis_Drain				: REFERENCE TO ST_Piston;
	stPis_CIP				: REFERENCE TO ST_Piston;
	
	stPis_Outlet: ST_Piston;
	tonDrainTime: TON;
	rt_Req_Reset: R_TRIG;
END_VAR

act_GetReference();

act_Oper();
//IF NOT Init.x THEN
	act_Status();
//END_IF

tonDrainTime(PT:=T#1M, IN:=eStatus=E_Line_Target.eDrain AND eReq=E_Line_Target.eNone);
IF tonDrainTime.Q 
AND eReq=E_Line_Target.eNone
AND eProcess=E_Line_Target.eNone
THEN;
	eReq:=E_Line_Target.eClose;
END_IF

m_Request_Reset(memo:=rt_Req_Reset);//

ACTION _aCIP_active:
bStepDone:=FALSE;
IF TRUE 
AND eStatus=E_Line_Target.eCIP
THEN;
	bStepDone:=TRUE;
END_IF
END_ACTION

ACTION _aCIP_entry:
fbPis.m_SetByRecipe(stPis:=stPis_TankA, 			req:=E_Piston_Recipe_State.Release);
//fbPis.m_SetByRecipe(stPis:=stPis_TankA_Pipe, 		req:=E_Piston_Recipe_State.Release);		
fbPis.m_SetByRecipe(stPis:=stPis_TankB, 			req:=E_Piston_Recipe_State.Release);
//fbPis.m_SetByRecipe(stPis:=stPis_TankB_Pipe, 		req:=E_Piston_Recipe_State.Release);
fbPis.m_SetByRecipe(stPis:=stPis_Drain, 			req:=E_Piston_Recipe_State.Act);
fbPis.m_SetByRecipe(stPis:=stPis_CIP, 				req:=E_Piston_Recipe_State.Act);
END_ACTION

ACTION _aClose_active:
bStepDone:=FALSE;
IF TRUE 
AND eStatus=E_Line_Target.eClose
THEN;
	bStepDone:=TRUE;
END_IF
END_ACTION

ACTION _aClose_entry:
fbPis.m_SetByRecipe(stPis:=stPis_TankA, 			req:=E_Piston_Recipe_State.Release);
//fbPis.m_SetByRecipe(stPis:=stPis_TankA_Pipe, 		req:=E_Piston_Recipe_State.Release);		
fbPis.m_SetByRecipe(stPis:=stPis_TankB, 			req:=E_Piston_Recipe_State.Release);
//fbPis.m_SetByRecipe(stPis:=stPis_TankB_Pipe, 		req:=E_Piston_Recipe_State.Release);
fbPis.m_SetByRecipe(stPis:=stPis_Drain, 			req:=E_Piston_Recipe_State.Release);
fbPis.m_SetByRecipe(stPis:=stPis_CIP, 				req:=E_Piston_Recipe_State.Release);
END_ACTION

ACTION _aDone_entry:
eProcess:=E_Line_Target.eNone;
eReq:=E_Line_Target.eNone;
bRun:=FALSE;
bDone:=TRUE;
END_ACTION

ACTION _aDrain_active:
bStepDone:=FALSE;
IF TRUE 
AND eStatus=E_Line_Target.eDrain
THEN;
	bStepDone:=TRUE;
END_IF
END_ACTION

ACTION _aDrain_entry:
fbPis.m_SetByRecipe(stPis:=stPis_TankA, 			req:=E_Piston_Recipe_State.Release);	
//fbPis.m_SetByRecipe(stPis:=stPis_TankA_Pipe, 		req:=E_Piston_Recipe_State.Release);	
fbPis.m_SetByRecipe(stPis:=stPis_TankB, 			req:=E_Piston_Recipe_State.Release);
//fbPis.m_SetByRecipe(stPis:=stPis_TankB_Pipe, 		req:=E_Piston_Recipe_State.Release);
fbPis.m_SetByRecipe(stPis:=stPis_Drain, 			req:=E_Piston_Recipe_State.Act);
fbPis.m_SetByRecipe(stPis:=stPis_CIP, 				req:=E_Piston_Recipe_State.Release);
END_ACTION

ACTION _aInit_active:
SFCReset:=FALSE;
END_ACTION

ACTION _aInit_exit:
eProcess:=E_Line_Target.eNone;
eReq:=E_Line_Target.eNone;
END_ACTION

ACTION _aReady_active:
CASE eReq OF
	E_Line_Target.eClose:;
			IF TRUE THEN;
				eProcess:=E_Line_Target.eClose;
			END_IF

	E_Line_Target.eTank_A:;
			IF TRUE THEN;
				eProcess:=E_Line_Target.eTank_A;
			END_IF	
			
	E_Line_Target.eTank_B:;
			IF TRUE THEN;
				eProcess:=E_Line_Target.eTank_B;
			END_IF	
			
	E_Line_Target.eCIP:;
			IF TRUE THEN;
				eProcess:=E_Line_Target.eCIP;
			END_IF	

	E_Line_Target.eDrain:;
			IF TRUE THEN;
				eProcess:=E_Line_Target.eDrain;
			END_IF	
		
END_CASE
END_ACTION

ACTION _aReady_exit:
bRun:=TRUE;
bDone:=FALSE;
END_ACTION

ACTION _aTank_A_active:
bStepDone:=FALSE;
IF TRUE  
AND eStatus=E_Line_Target.eTank_A 
THEN;
	bStepDone:=TRUE;
END_IF
END_ACTION

ACTION _aTank_A_entry:
fbPis.m_SetByRecipe(stPis:=stPis_TankA, 			req:=E_Piston_Recipe_State.Act);	
fbPis.m_SetByRecipe(stPis:=stPis_TankA_Pipe, 		req:=E_Piston_Recipe_State.Release);	
fbPis.m_SetByRecipe(stPis:=stPis_TankB, 			req:=E_Piston_Recipe_State.Release);
//fbPis.m_SetByRecipe(stPis:=stPis_TankB_Pipe, 		req:=E_Piston_Recipe_State.Release);
fbPis.m_SetByRecipe(stPis:=stPis_Drain, 			req:=E_Piston_Recipe_State.Release);
fbPis.m_SetByRecipe(stPis:=stPis_CIP, 				req:=E_Piston_Recipe_State.Release);
END_ACTION

ACTION _aTank_B_active:
bStepDone:=FALSE;
IF TRUE 
AND eStatus=E_Line_Target.eTank_B
THEN;
	bStepDone:=TRUE;
END_IF
END_ACTION

ACTION _aTank_B_entry:
fbPis.m_SetByRecipe(stPis:=stPis_TankA, 			req:=E_Piston_Recipe_State.Release);	
//fbPis.m_SetByRecipe(stPis:=stPis_TankA_Pipe, 		req:=E_Piston_Recipe_State.Release);	
fbPis.m_SetByRecipe(stPis:=stPis_TankB, 			req:=E_Piston_Recipe_State.Act);
fbPis.m_SetByRecipe(stPis:=stPis_TankB_Pipe, 		req:=E_Piston_Recipe_State.Release);
fbPis.m_SetByRecipe(stPis:=stPis_Drain, 			req:=E_Piston_Recipe_State.Release);
fbPis.m_SetByRecipe(stPis:=stPis_CIP, 				req:=E_Piston_Recipe_State.Release);
END_ACTION

ACTION act_GetReference:
m_Set_SFCFlags_Reference();
//refElement REF= fbElement[eElementID];
//refState_Long REF= fbElement[eElementID].eState_Long;

stPis_TankA				REF= g_Piston.stPis[valTankA];
stPis_TankB				REF= g_Piston.stPis[valTankB];
stPis_TankA_Pipe		REF= g_Piston.stPis[valTankA_Pipe];
stPis_TankB_Pipe		REF= g_Piston.stPis[valTankB_Pipe];
stPis_Drain				REF= g_Piston.stPis[valDrain];
stPis_CIP				REF= g_Piston.stPis[valCIP];
END_ACTION

ACTION act_Oper:
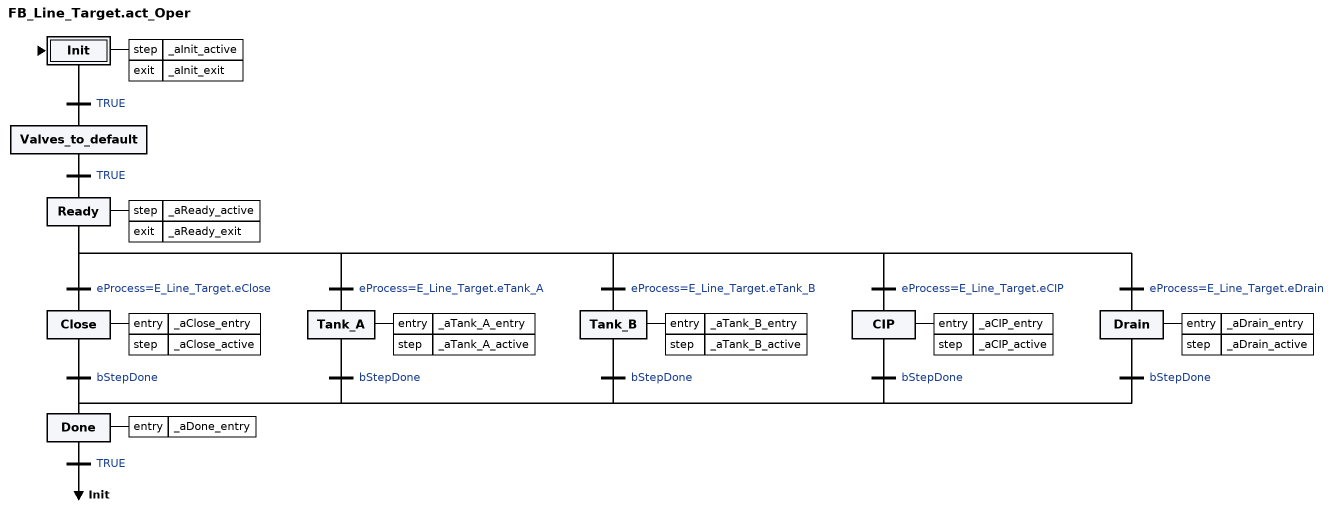
INITIAL_STEP Init:
    _aInit_active(N);  // step action
    _aInit_exit(P0);  // exit action
END_STEP
TRANSITION FROM Init TO Valves_to_default
    := TRUE;
END_TRANSITION
STEP Valves_to_default:
END_STEP
TRANSITION FROM Valves_to_default TO Ready
    := TRUE;
END_TRANSITION
STEP Ready:
    _aReady_active(N);  // step action
    _aReady_exit(P0);  // exit action
END_STEP
TRANSITION FROM Ready TO Close
    := eProcess=E_Line_Target.eClose;
END_TRANSITION
STEP Close:  // min time t#1s
    _aClose_entry(P1);  // entry action
    _aClose_active(N);  // step action
END_STEP
TRANSITION FROM Close TO Done
    := bStepDone;
END_TRANSITION
TRANSITION FROM Ready TO Tank_A
    := eProcess=E_Line_Target.eTank_A;
END_TRANSITION
STEP Tank_A:  // min time t#1s
    _aTank_A_entry(P1);  // entry action
    _aTank_A_active(N);  // step action
END_STEP
TRANSITION FROM Tank_A TO Done
    := bStepDone;
END_TRANSITION
TRANSITION FROM Ready TO Tank_B
    := eProcess=E_Line_Target.eTank_B;
END_TRANSITION
STEP Tank_B:  // min time t#1s
    _aTank_B_entry(P1);  // entry action
    _aTank_B_active(N);  // step action
END_STEP
TRANSITION FROM Tank_B TO Done
    := bStepDone;
END_TRANSITION
TRANSITION FROM Ready TO CIP
    := eProcess=E_Line_Target.eCIP;
END_TRANSITION
STEP CIP:  // min time t#1s
    _aCIP_entry(P1);  // entry action
    _aCIP_active(N);  // step action
END_STEP
TRANSITION FROM CIP TO Done
    := bStepDone;
END_TRANSITION
TRANSITION FROM Ready TO Drain
    := eProcess=E_Line_Target.eDrain;
END_TRANSITION
STEP Drain:  // min time t#1s
    _aDrain_entry(P1);  // entry action
    _aDrain_active(N);  // step action
END_STEP
TRANSITION FROM Drain TO Done
    := bStepDone;
END_TRANSITION
STEP Done:
    _aDone_entry(P1);  // entry action
END_STEP
TRANSITION FROM Done TO Init
    := TRUE;
END_TRANSITION
// branch label Branch0_act_Oper
END_ACTION

